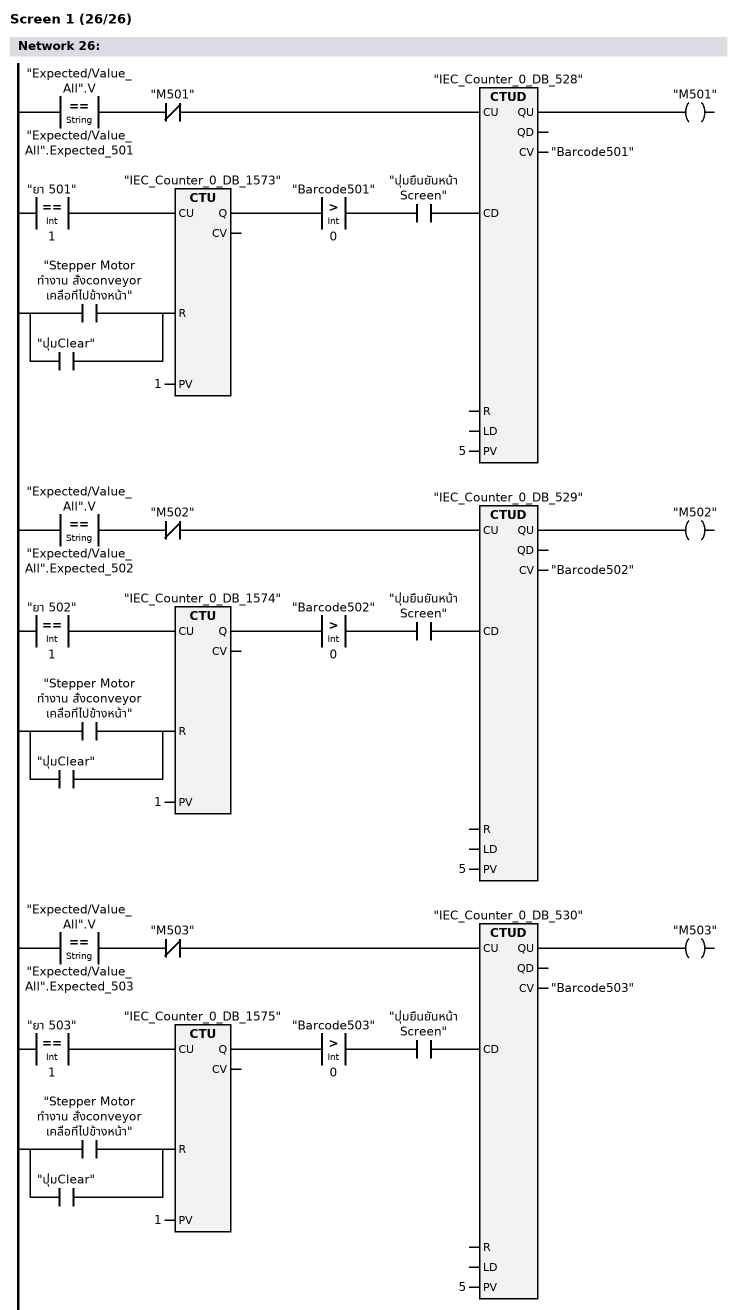
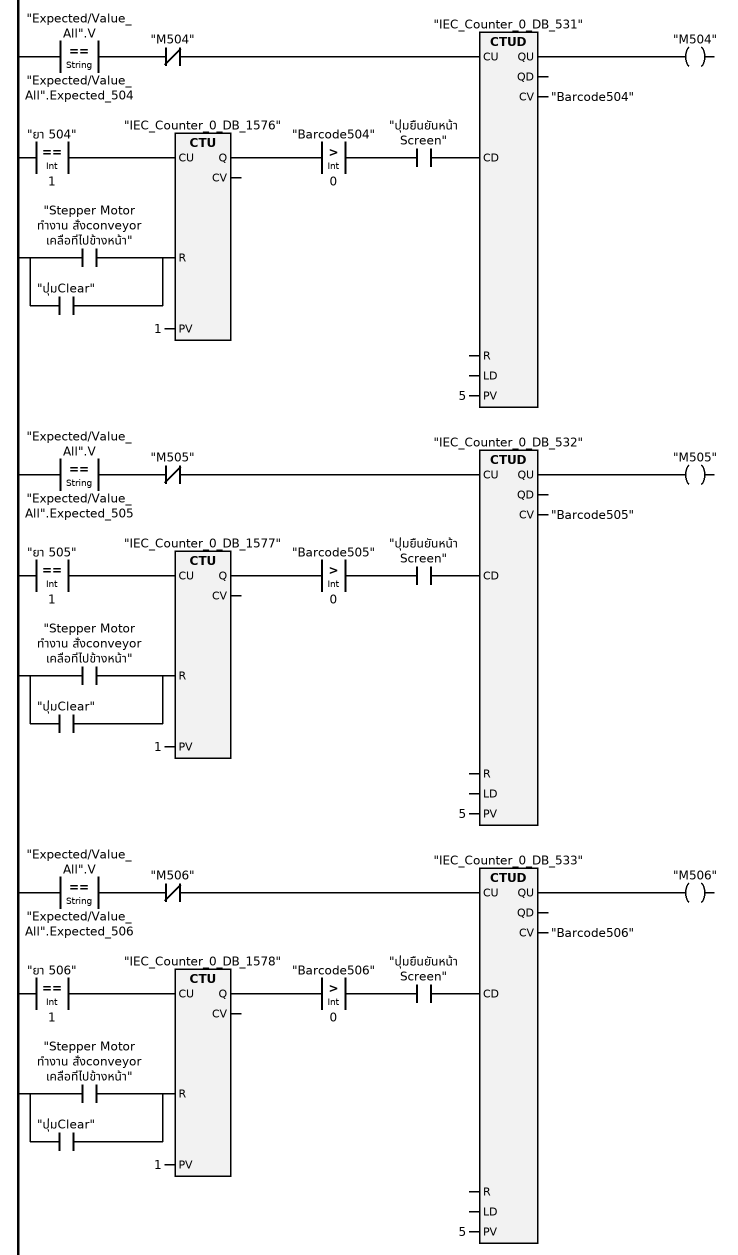
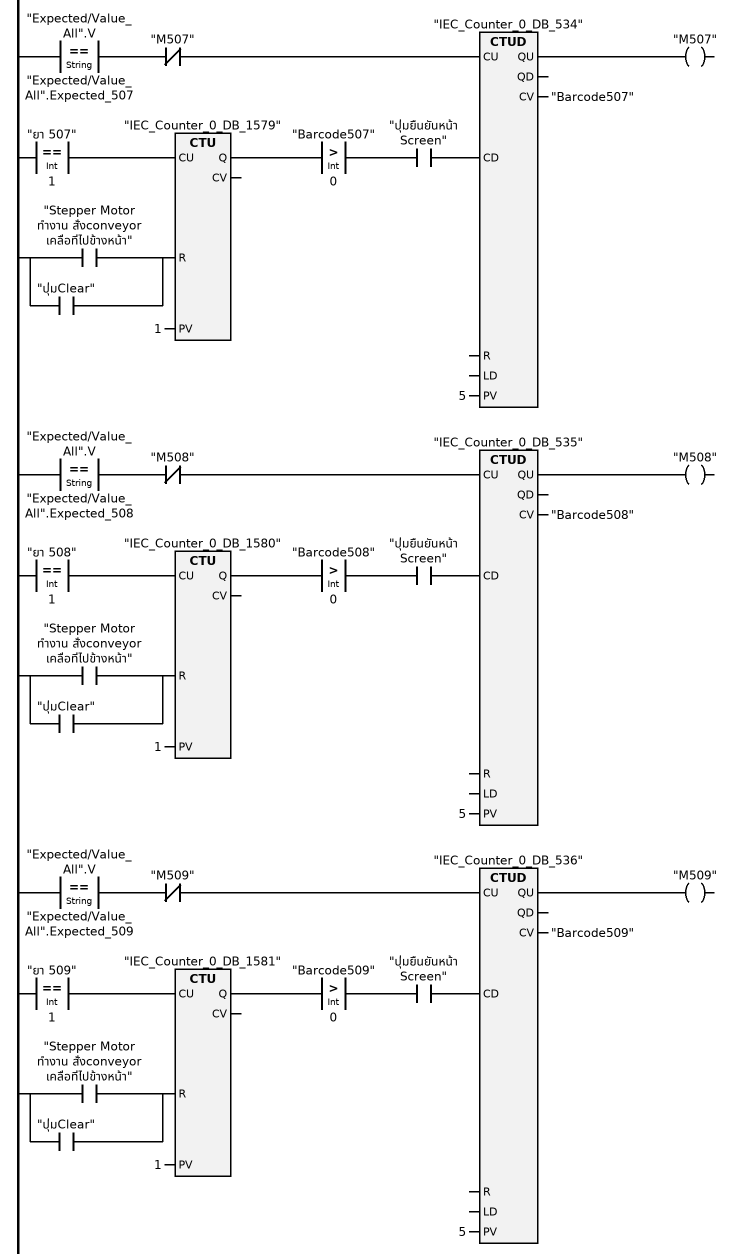
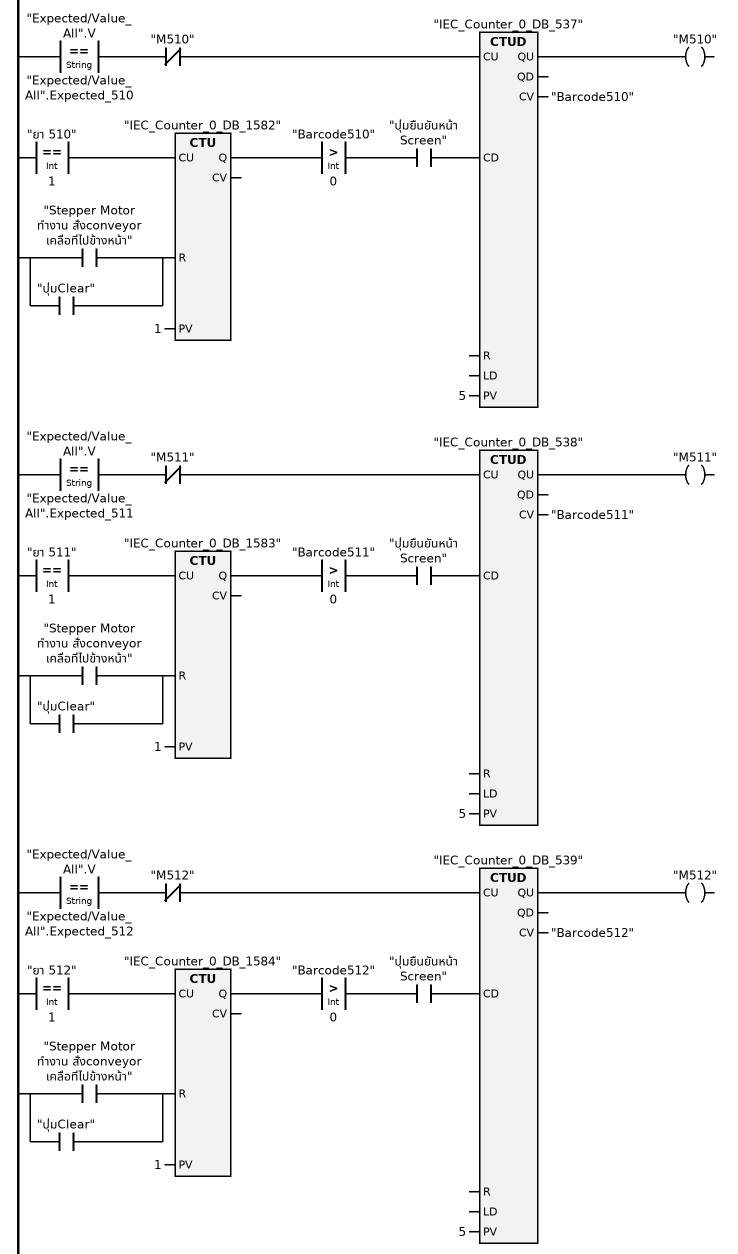
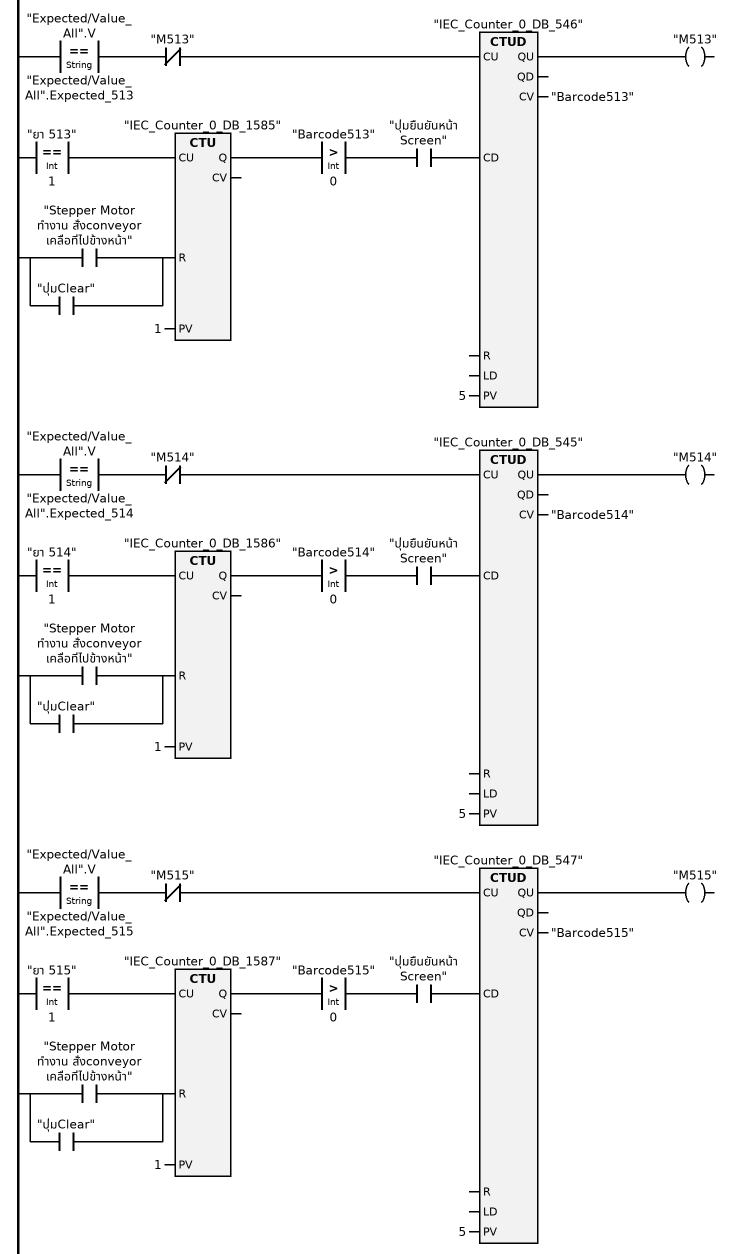
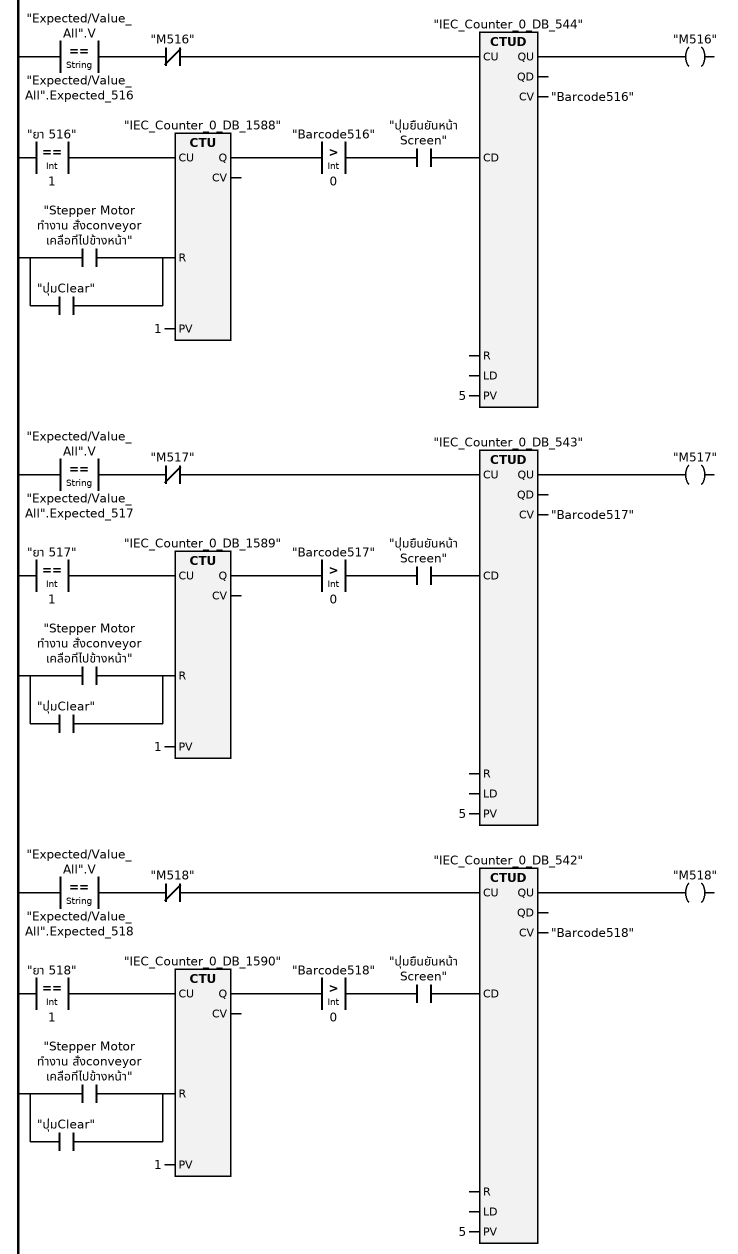
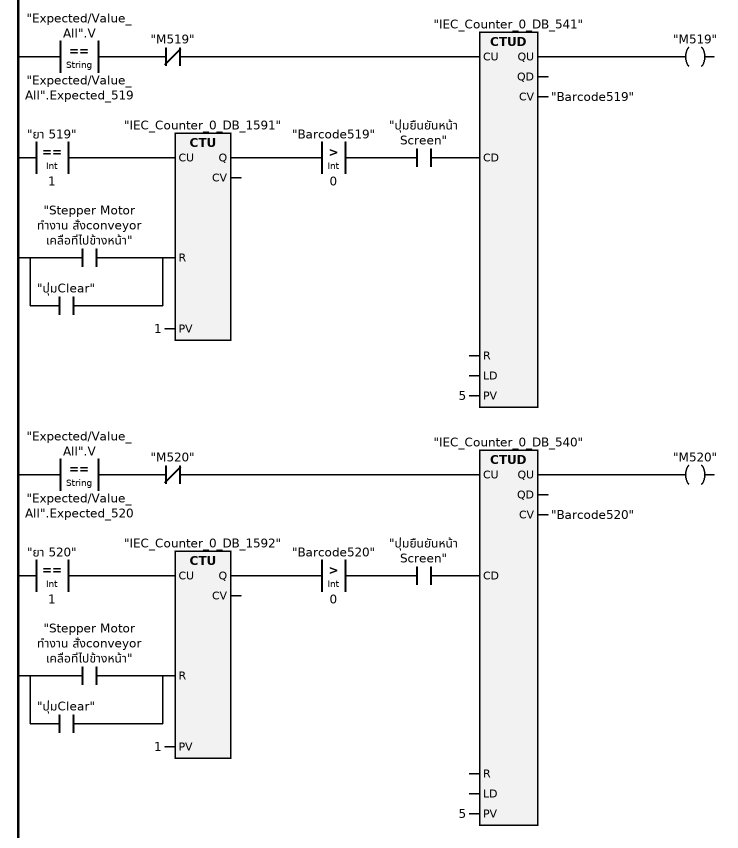
   "IEC_Counter_0_DB_1573".CTU(CU := "ยา 501" = 1,
                           R := "Stepper Motor ทำงาน สั่งconveyor เคลื่อที่ไปข้างหน้า" OR "ปุ่มClear",
                           PV := 1);
   "IEC_Counter_0_DB_528".CTUD(CU := ("Expected/Value_All".V = "Expected/Value_All".Expected_501) AND NOT "M501",
                           CD := "IEC_Counter_0_DB_1573".Q AND ("Barcode501" > 0) AND "ปุ่มยืนยันหน้า Screen",
                           PV := 5,
                           CV => "Barcode501");
   "M501" := "IEC_Counter_0_DB_528".QU;
   "IEC_Counter_0_DB_1574".CTU(CU := "ยา 502" = 1,
                           R := "Stepper Motor ทำงาน สั่งconveyor เคลื่อที่ไปข้างหน้า" OR "ปุ่มClear",
                           PV := 1);
   "IEC_Counter_0_DB_529".CTUD(CU := ("Expected/Value_All".V = "Expected/Value_All".Expected_502) AND NOT "M502",
                           CD := "IEC_Counter_0_DB_1574".Q AND ("Barcode502" > 0) AND "ปุ่มยืนยันหน้า Screen",
                           PV := 5,
                           CV => "Barcode502");
   "M502" := "IEC_Counter_0_DB_529".QU;
   "IEC_Counter_0_DB_1575".CTU(CU := "ยา 503" = 1,
                           R := "Stepper Motor ทำงาน สั่งconveyor เคลื่อที่ไปข้างหน้า" OR "ปุ่มClear",
                           PV := 1);
   "IEC_Counter_0_DB_530".CTUD(CU := ("Expected/Value_All".V = "Expected/Value_All".Expected_503) AND NOT "M503",
                           CD := "IEC_Counter_0_DB_1575".Q AND ("Barcode503" > 0) AND "ปุ่มยืนยันหน้า Screen",
                           PV := 5,
                           CV => "Barcode503");
   "M503" := "IEC_Counter_0_DB_530".QU;
   "IEC_Counter_0_DB_1576".CTU(CU := "ยา 504" = 1,
                           R := "Stepper Motor ทำงาน สั่งconveyor เคลื่อที่ไปข้างหน้า" OR "ปุ่มClear",
                           PV := 1);
   "IEC_Counter_0_DB_531".CTUD(CU := ("Expected/Value_All".V = "Expected/Value_All".Expected_504) AND NOT "M504",
                           CD := "IEC_Counter_0_DB_1576".Q AND ("Barcode504" > 0) AND "ปุ่มยืนยันหน้า Screen",
                           PV := 5,
                           CV => "Barcode504");
   "M504" := "IEC_Counter_0_DB_531".QU;
   "IEC_Counter_0_DB_1577".CTU(CU := "ยา 505" = 1,
                           R := "Stepper Motor ทำงาน สั่งconveyor เคลื่อที่ไปข้างหน้า" OR "ปุ่มClear",
                           PV := 1);
   "IEC_Counter_0_DB_532".CTUD(CU := ("Expected/Value_All".V = "Expected/Value_All".Expected_505) AND NOT "M505",
                           CD := "IEC_Counter_0_DB_1577".Q AND ("Barcode505" > 0) AND "ปุ่มยืนยันหน้า Screen",
                           PV := 5,
                           CV => "Barcode505");
   "M505" := "IEC_Counter_0_DB_532".QU;
   "IEC_Counter_0_DB_1578".CTU(CU := "ยา 506" = 1,
                           R := "Stepper Motor ทำงาน สั่งconveyor เคลื่อที่ไปข้างหน้า" OR "ปุ่มClear",
                           PV := 1);
   "IEC_Counter_0_DB_533".CTUD(CU := ("Expected/Value_All".V = "Expected/Value_All".Expected_506) AND NOT "M506",
                           CD := "IEC_Counter_0_DB_1578".Q AND ("Barcode506" > 0) AND "ปุ่มยืนยันหน้า Screen",
                           PV := 5,
                           CV => "Barcode506");
   "M506" := "IEC_Counter_0_DB_533".QU;
   "IEC_Counter_0_DB_1579".CTU(CU := "ยา 507" = 1,
                           R := "Stepper Motor ทำงาน สั่งconveyor เคลื่อที่ไปข้างหน้า" OR "ปุ่มClear",
                           PV := 1);
   "IEC_Counter_0_DB_534".CTUD(CU := ("Expected/Value_All".V = "Expected/Value_All".Expected_507) AND NOT "M507",
                           CD := "IEC_Counter_0_DB_1579".Q AND ("Barcode507" > 0) AND "ปุ่มยืนยันหน้า Screen",
                           PV := 5,
                           CV => "Barcode507");
   "M507" := "IEC_Counter_0_DB_534".QU;
   "IEC_Counter_0_DB_1580".CTU(CU := "ยา 508" = 1,
                           R := "Stepper Motor ทำงาน สั่งconveyor เคลื่อที่ไปข้างหน้า" OR "ปุ่มClear",
                           PV := 1);
   "IEC_Counter_0_DB_535".CTUD(CU := ("Expected/Value_All".V = "Expected/Value_All".Expected_508) AND NOT "M508",
                           CD := "IEC_Counter_0_DB_1580".Q AND ("Barcode508" > 0) AND "ปุ่มยืนยันหน้า Screen",
                           PV := 5,
                           CV => "Barcode508");
   "M508" := "IEC_Counter_0_DB_535".QU;
   "IEC_Counter_0_DB_1581".CTU(CU := "ยา 509" = 1,
                           R := "Stepper Motor ทำงาน สั่งconveyor เคลื่อที่ไปข้างหน้า" OR "ปุ่มClear",
                           PV := 1);
   "IEC_Counter_0_DB_536".CTUD(CU := ("Expected/Value_All".V = "Expected/Value_All".Expected_509) AND NOT "M509",
                           CD := "IEC_Counter_0_DB_1581".Q AND ("Barcode509" > 0) AND "ปุ่มยืนยันหน้า Screen",
                           PV := 5,
                           CV => "Barcode509");
   "M509" := "IEC_Counter_0_DB_536".QU;
   "IEC_Counter_0_DB_1582".CTU(CU := "ยา 510" = 1,
                           R := "Stepper Motor ทำงาน สั่งconveyor เคลื่อที่ไปข้างหน้า" OR "ปุ่มClear",
                           PV := 1);
   "IEC_Counter_0_DB_537".CTUD(CU := ("Expected/Value_All".V = "Expected/Value_All".Expected_510) AND NOT "M510",
                           CD := "IEC_Counter_0_DB_1582".Q AND ("Barcode510" > 0) AND "ปุ่มยืนยันหน้า Screen",
                           PV := 5,
                           CV => "Barcode510");
   "M510" := "IEC_Counter_0_DB_537".QU;
   "IEC_Counter_0_DB_1583".CTU(CU := "ยา 511" = 1,
                           R := "Stepper Motor ทำงาน สั่งconveyor เคลื่อที่ไปข้างหน้า" OR "ปุ่มClear",
                           PV := 1);
   "IEC_Counter_0_DB_538".CTUD(CU := ("Expected/Value_All".V = "Expected/Value_All".Expected_511) AND NOT "M511",
                           CD := "IEC_Counter_0_DB_1583".Q AND ("Barcode511" > 0) AND "ปุ่มยืนยันหน้า Screen",
                           PV := 5,
                           CV => "Barcode511");
   "M511" := "IEC_Counter_0_DB_538".QU;
   "IEC_Counter_0_DB_1584".CTU(CU := "ยา 512" = 1,
                           R := "Stepper Motor ทำงาน สั่งconveyor เคลื่อที่ไปข้างหน้า" OR "ปุ่มClear",
                           PV := 1);
   "IEC_Counter_0_DB_539".CTUD(CU := ("Expected/Value_All".V = "Expected/Value_All".Expected_512) AND NOT "M512",
                           CD := "IEC_Counter_0_DB_1584".Q AND ("Barcode512" > 0) AND "ปุ่มยืนยันหน้า Screen",
                           PV := 5,
                           CV => "Barcode512");
   "M512" := "IEC_Counter_0_DB_539".QU;
   "IEC_Counter_0_DB_1585".CTU(CU := "ยา 513" = 1,
                           R := "Stepper Motor ทำงาน สั่งconveyor เคลื่อที่ไปข้างหน้า" OR "ปุ่มClear",
                           PV := 1);
   "IEC_Counter_0_DB_546".CTUD(CU := ("Expected/Value_All".V = "Expected/Value_All".Expected_513) AND NOT "M513",
                           CD := "IEC_Counter_0_DB_1585".Q AND ("Barcode513" > 0) AND "ปุ่มยืนยันหน้า Screen",
                           PV := 5,
                           CV => "Barcode513");
   "M513" := "IEC_Counter_0_DB_546".QU;
   "IEC_Counter_0_DB_1586".CTU(CU := "ยา 514" = 1,
                           R := "Stepper Motor ทำงาน สั่งconveyor เคลื่อที่ไปข้างหน้า" OR "ปุ่มClear",
                           PV := 1);
   "IEC_Counter_0_DB_545".CTUD(CU := ("Expected/Value_All".V = "Expected/Value_All".Expected_514) AND NOT "M514",
                           CD := "IEC_Counter_0_DB_1586".Q AND ("Barcode514" > 0) AND "ปุ่มยืนยันหน้า Screen",
                           PV := 5,
                           CV => "Barcode514");
   "M514" := "IEC_Counter_0_DB_545".QU;
   "IEC_Counter_0_DB_1587".CTU(CU := "ยา 515" = 1,
                           R := "Stepper Motor ทำงาน สั่งconveyor เคลื่อที่ไปข้างหน้า" OR "ปุ่มClear",
                           PV := 1);
   "IEC_Counter_0_DB_547".CTUD(CU := ("Expected/Value_All".V = "Expected/Value_All".Expected_515) AND NOT "M515",
                           CD := "IEC_Counter_0_DB_1587".Q AND ("Barcode515" > 0) AND "ปุ่มยืนยันหน้า Screen",
                           PV := 5,
                           CV => "Barcode515");
   "M515" := "IEC_Counter_0_DB_547".QU;
   "IEC_Counter_0_DB_1588".CTU(CU := "ยา 516" = 1,
                           R := "Stepper Motor ทำงาน สั่งconveyor เคลื่อที่ไปข้างหน้า" OR "ปุ่มClear",
                           PV := 1);
   "IEC_Counter_0_DB_544".CTUD(CU := ("Expected/Value_All".V = "Expected/Value_All".Expected_516) AND NOT "M516",
                           CD := "IEC_Counter_0_DB_1588".Q AND ("Barcode516" > 0) AND "ปุ่มยืนยันหน้า Screen",
                           PV := 5,
                           CV => "Barcode516");
   "M516" := "IEC_Counter_0_DB_544".QU;
   "IEC_Counter_0_DB_1589".CTU(CU := "ยา 517" = 1,
                           R := "Stepper Motor ทำงาน สั่งconveyor เคลื่อที่ไปข้างหน้า" OR "ปุ่มClear",
                           PV := 1);
   "IEC_Counter_0_DB_543".CTUD(CU := ("Expected/Value_All".V = "Expected/Value_All".Expected_517) AND NOT "M517",
                           CD := "IEC_Counter_0_DB_1589".Q AND ("Barcode517" > 0) AND "ปุ่มยืนยันหน้า Screen",
                           PV := 5,
                           CV => "Barcode517");
   "M517" := "IEC_Counter_0_DB_543".QU;
   "IEC_Counter_0_DB_1590".CTU(CU := "ยา 518" = 1,
                           R := "Stepper Motor ทำงาน สั่งconveyor เคลื่อที่ไปข้างหน้า" OR "ปุ่มClear",
                           PV := 1);
   "IEC_Counter_0_DB_542".CTUD(CU := ("Expected/Value_All".V = "Expected/Value_All".Expected_518) AND NOT "M518",
                           CD := "IEC_Counter_0_DB_1590".Q AND ("Barcode518" > 0) AND "ปุ่มยืนยันหน้า Screen",
                           PV := 5,
                           CV => "Barcode518");
   "M518" := "IEC_Counter_0_DB_542".QU;
   "IEC_Counter_0_DB_1591".CTU(CU := "ยา 519" = 1,
                           R := "Stepper Motor ทำงาน สั่งconveyor เคลื่อที่ไปข้างหน้า" OR "ปุ่มClear",
                           PV := 1);
   "IEC_Counter_0_DB_541".CTUD(CU := ("Expected/Value_All".V = "Expected/Value_All".Expected_519) AND NOT "M519",
                           CD := "IEC_Counter_0_DB_1591".Q AND ("Barcode519" > 0) AND "ปุ่มยืนยันหน้า Screen",
                           PV := 5,
                           CV => "Barcode519");
   "M519" := "IEC_Counter_0_DB_541".QU;
   "IEC_Counter_0_DB_1592".CTU(CU := "ยา 520" = 1,
                           R := "Stepper Motor ทำงาน สั่งconveyor เคลื่อที่ไปข้างหน้า" OR "ปุ่มClear",
                           PV := 1);
   "IEC_Counter_0_DB_540".CTUD(CU := ("Expected/Value_All".V = "Expected/Value_All".Expected_520) AND NOT "M520",
                           CD := "IEC_Counter_0_DB_1592".Q AND ("Barcode520" > 0) AND "ปุ่มยืนยันหน้า Screen",
                           PV := 5,
                           CV => "Barcode520");
   "M520" := "IEC_Counter_0_DB_540".QU;
END_REGION
END_FUNCTION

FUNCTION "Screen2" : Void   // FC14, LAD
{ S7_Optimized_Access := 'TRUE' }
VERSION : 0.1
   VAR_OUTPUT
      Output : Word;
   END_VAR
BEGIN

REGION Network 1
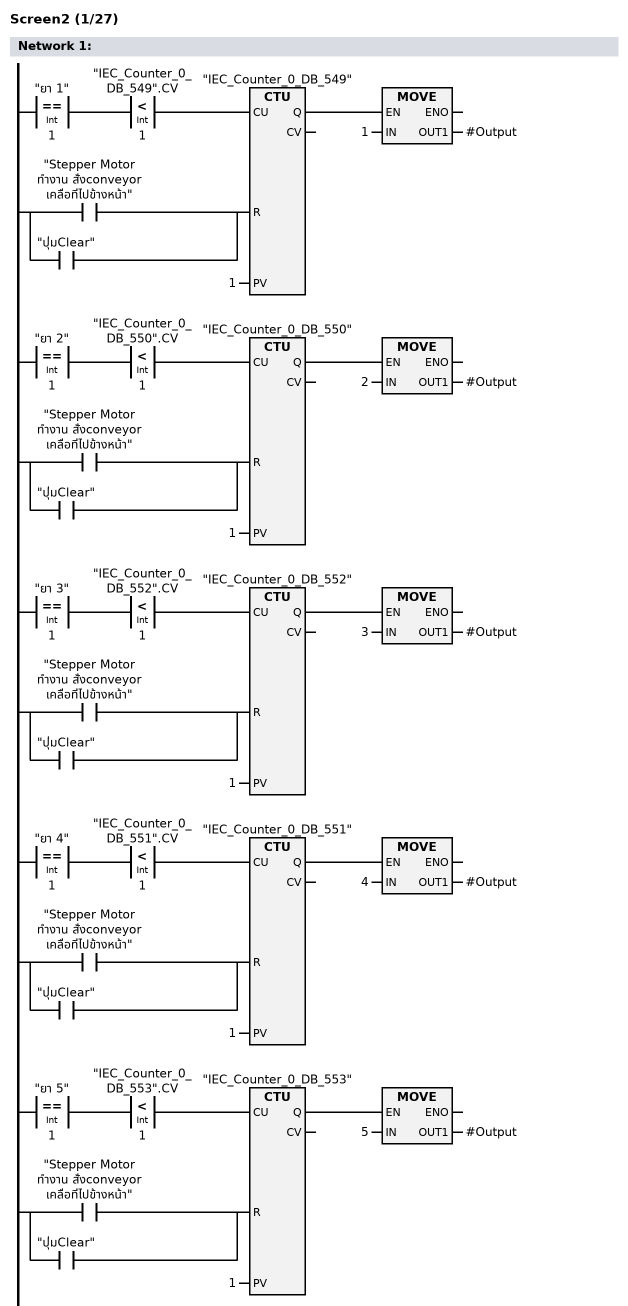
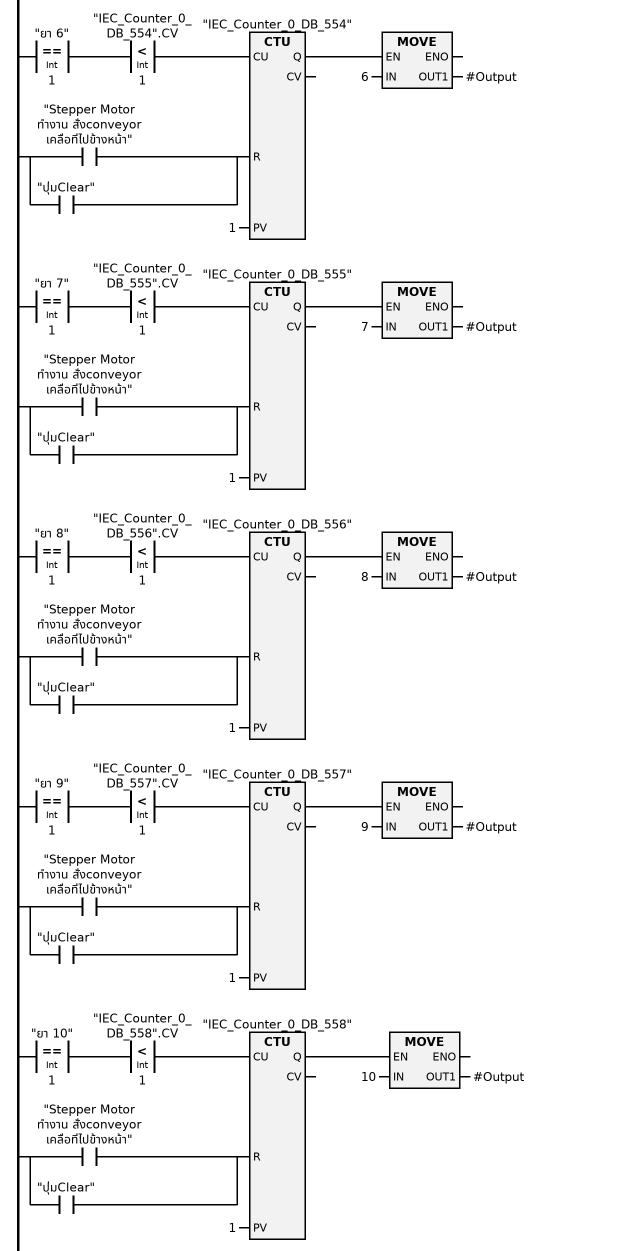
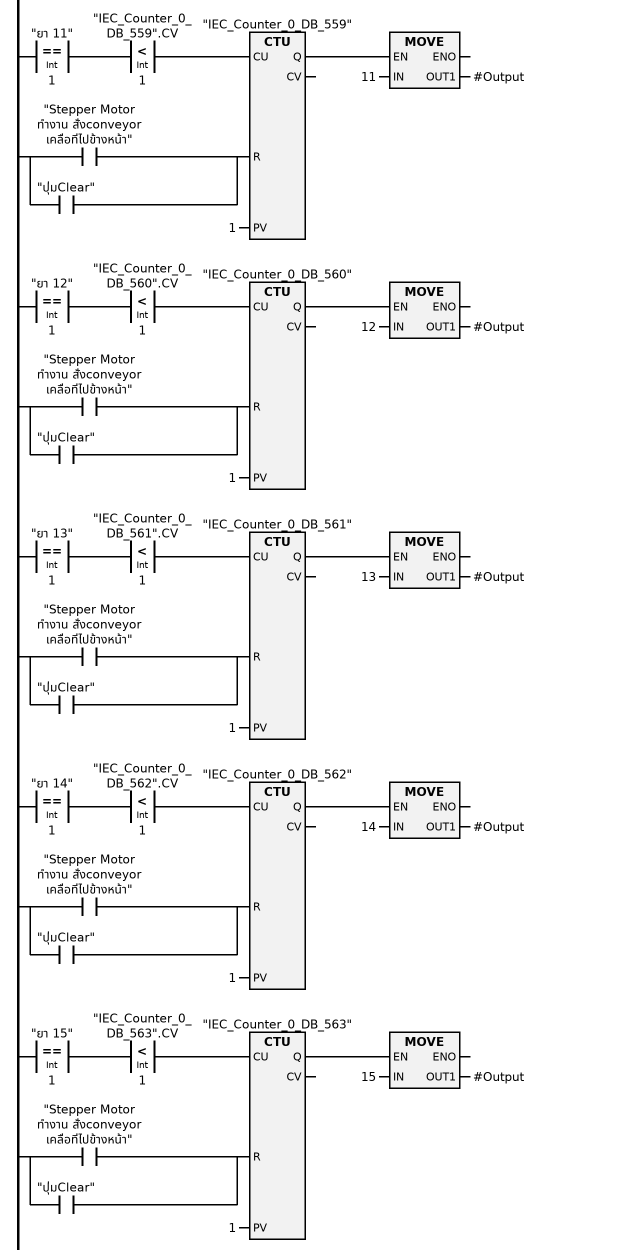
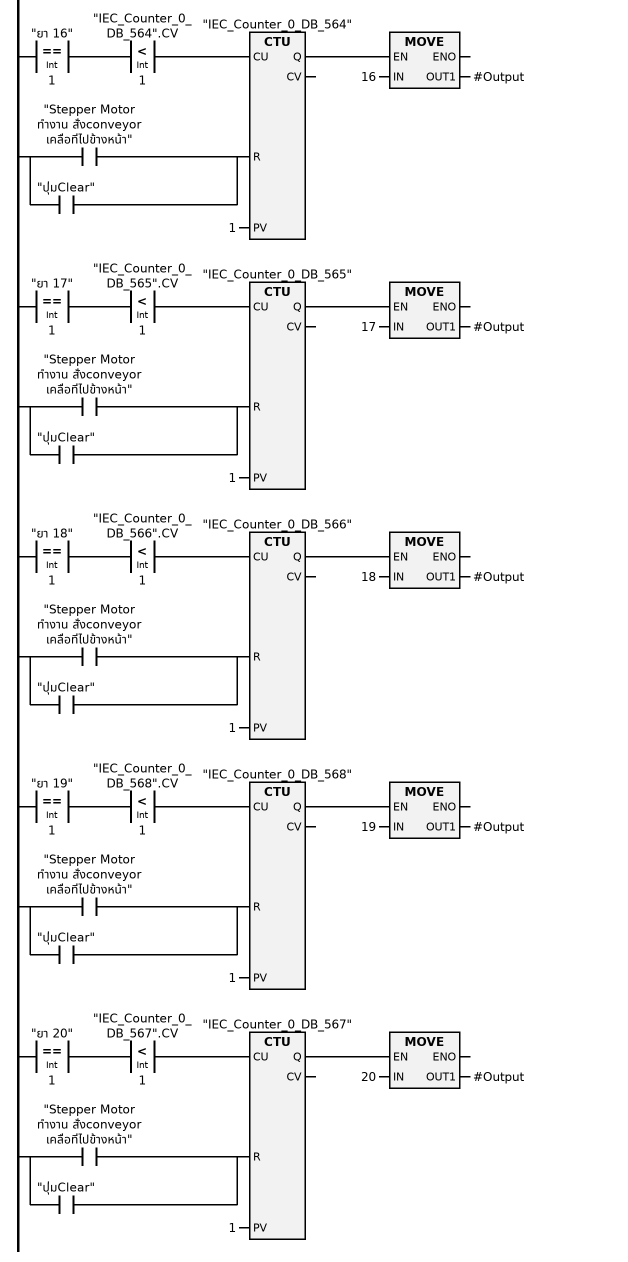
   "IEC_Counter_0_DB_549".CTU(CU := ("ยา 1" = 1) AND ("IEC_Counter_0_DB_549".CV < 1),
                           R := "Stepper Motor ทำงาน สั่งconveyor เคลื่อที่ไปข้างหน้า" OR "ปุ่มClear",
                           PV := 1);
   IF "IEC_Counter_0_DB_549".Q THEN #Output := 1; END_IF;
   "IEC_Counter_0_DB_550".CTU(CU := ("ยา 2" = 1) AND ("IEC_Counter_0_DB_550".CV < 1),
                           R := "Stepper Motor ทำงาน สั่งconveyor เคลื่อที่ไปข้างหน้า" OR "ปุ่มClear",
                           PV := 1);
   IF "IEC_Counter_0_DB_550".Q THEN #Output := 2; END_IF;
   "IEC_Counter_0_DB_552".CTU(CU := ("ยา 3" = 1) AND ("IEC_Counter_0_DB_552".CV < 1),
                           R := "Stepper Motor ทำงาน สั่งconveyor เคลื่อที่ไปข้างหน้า" OR "ปุ่มClear",
                           PV := 1);
   IF "IEC_Counter_0_DB_552".Q THEN #Output := 3; END_IF;
   "IEC_Counter_0_DB_551".CTU(CU := ("ยา 4" = 1) AND ("IEC_Counter_0_DB_551".CV < 1),
                           R := "Stepper Motor ทำงาน สั่งconveyor เคลื่อที่ไปข้างหน้า" OR "ปุ่มClear",
                           PV := 1);
   IF "IEC_Counter_0_DB_551".Q THEN #Output := 4; END_IF;
   "IEC_Counter_0_DB_553".CTU(CU := ("ยา 5" = 1) AND ("IEC_Counter_0_DB_553".CV < 1),
                           R := "Stepper Motor ทำงาน สั่งconveyor เคลื่อที่ไปข้างหน้า" OR "ปุ่มClear",
                           PV := 1);
   IF "IEC_Counter_0_DB_553".Q THEN #Output := 5; END_IF;
   "IEC_Counter_0_DB_554".CTU(CU := ("ยา 6" = 1) AND ("IEC_Counter_0_DB_554".CV < 1),
                           R := "Stepper Motor ทำงาน สั่งconveyor เคลื่อที่ไปข้างหน้า" OR "ปุ่มClear",
                           PV := 1);
   IF "IEC_Counter_0_DB_554".Q THEN #Output := 6; END_IF;
   "IEC_Counter_0_DB_555".CTU(CU := ("ยา 7" = 1) AND ("IEC_Counter_0_DB_555".CV < 1),
                           R := "Stepper Motor ทำงาน สั่งconveyor เคลื่อที่ไปข้างหน้า" OR "ปุ่มClear",
                           PV := 1);
   IF "IEC_Counter_0_DB_555".Q THEN #Output := 7; END_IF;
   "IEC_Counter_0_DB_556".CTU(CU := ("ยา 8" = 1) AND ("IEC_Counter_0_DB_556".CV < 1),
                           R := "Stepper Motor ทำงาน สั่งconveyor เคลื่อที่ไปข้างหน้า" OR "ปุ่มClear",
                           PV := 1);
   IF "IEC_Counter_0_DB_556".Q THEN #Output := 8; END_IF;
   "IEC_Counter_0_DB_557".CTU(CU := ("ยา 9" = 1) AND ("IEC_Counter_0_DB_557".CV < 1),
                           R := "Stepper Motor ทำงาน สั่งconveyor เคลื่อที่ไปข้างหน้า" OR "ปุ่มClear",
                           PV := 1);
   IF "IEC_Counter_0_DB_557".Q THEN #Output := 9; END_IF;
   "IEC_Counter_0_DB_558".CTU(CU := ("ยา 10" = 1) AND ("IEC_Counter_0_DB_558".CV < 1),
                           R := "Stepper Motor ทำงาน สั่งconveyor เคลื่อที่ไปข้างหน้า" OR "ปุ่มClear",
                           PV := 1);
   IF "IEC_Counter_0_DB_558".Q THEN #Output := 10; END_IF;
   "IEC_Counter_0_DB_559".CTU(CU := ("ยา 11" = 1) AND ("IEC_Counter_0_DB_559".CV < 1),
                           R := "Stepper Motor ทำงาน สั่งconveyor เคลื่อที่ไปข้างหน้า" OR "ปุ่มClear",
                           PV := 1);
   IF "IEC_Counter_0_DB_559".Q THEN #Output := 11; END_IF;
   "IEC_Counter_0_DB_560".CTU(CU := ("ยา 12" = 1) AND ("IEC_Counter_0_DB_560".CV < 1),
                           R := "Stepper Motor ทำงาน สั่งconveyor เคลื่อที่ไปข้างหน้า" OR "ปุ่มClear",
                           PV := 1);
   IF "IEC_Counter_0_DB_560".Q THEN #Output := 12; END_IF;
   "IEC_Counter_0_DB_561".CTU(CU := ("ยา 13" = 1) AND ("IEC_Counter_0_DB_561".CV < 1),
                           R := "Stepper Motor ทำงาน สั่งconveyor เคลื่อที่ไปข้างหน้า" OR "ปุ่มClear",
                           PV := 1);
   IF "IEC_Counter_0_DB_561".Q THEN #Output := 13; END_IF;
   "IEC_Counter_0_DB_562".CTU(CU := ("ยา 14" = 1) AND ("IEC_Counter_0_DB_562".CV < 1),
                           R := "Stepper Motor ทำงาน สั่งconveyor เคลื่อที่ไปข้างหน้า" OR "ปุ่มClear",
                           PV := 1);
   IF "IEC_Counter_0_DB_562".Q THEN #Output := 14; END_IF;
   "IEC_Counter_0_DB_563".CTU(CU := ("ยา 15" = 1) AND ("IEC_Counter_0_DB_563".CV < 1),
                           R := "Stepper Motor ทำงาน สั่งconveyor เคลื่อที่ไปข้างหน้า" OR "ปุ่มClear",
                           PV := 1);
   IF "IEC_Counter_0_DB_563".Q THEN #Output := 15; END_IF;
   "IEC_Counter_0_DB_564".CTU(CU := ("ยา 16" = 1) AND ("IEC_Counter_0_DB_564".CV < 1),
                           R := "Stepper Motor ทำงาน สั่งconveyor เคลื่อที่ไปข้างหน้า" OR "ปุ่มClear",
                           PV := 1);
   IF "IEC_Counter_0_DB_564".Q THEN #Output := 16; END_IF;
   "IEC_Counter_0_DB_565".CTU(CU := ("ยา 17" = 1) AND ("IEC_Counter_0_DB_565".CV < 1),
                           R := "Stepper Motor ทำงาน สั่งconveyor เคลื่อที่ไปข้างหน้า" OR "ปุ่มClear",
                           PV := 1);
   IF "IEC_Counter_0_DB_565".Q THEN #Output := 17; END_IF;
   "IEC_Counter_0_DB_566".CTU(CU := ("ยา 18" = 1) AND ("IEC_Counter_0_DB_566".CV < 1),
                           R := "Stepper Motor ทำงาน สั่งconveyor เคลื่อที่ไปข้างหน้า" OR "ปุ่มClear",
                           PV := 1);
   IF "IEC_Counter_0_DB_566".Q THEN #Output := 18; END_IF;
   "IEC_Counter_0_DB_568".CTU(CU := ("ยา 19" = 1) AND ("IEC_Counter_0_DB_568".CV < 1),
                           R := "Stepper Motor ทำงาน สั่งconveyor เคลื่อที่ไปข้างหน้า" OR "ปุ่มClear",
                           PV := 1);
   IF "IEC_Counter_0_DB_568".Q THEN #Output := 19; END_IF;
   "IEC_Counter_0_DB_567".CTU(CU := ("ยา 20" = 1) AND ("IEC_Counter_0_DB_567".CV < 1),
                           R := "Stepper Motor ทำงาน สั่งconveyor เคลื่อที่ไปข้างหน้า" OR "ปุ่มClear",
                           PV := 1);
   IF "IEC_Counter_0_DB_567".Q THEN #Output := 20; END_IF;
END_REGION

REGION Network 2
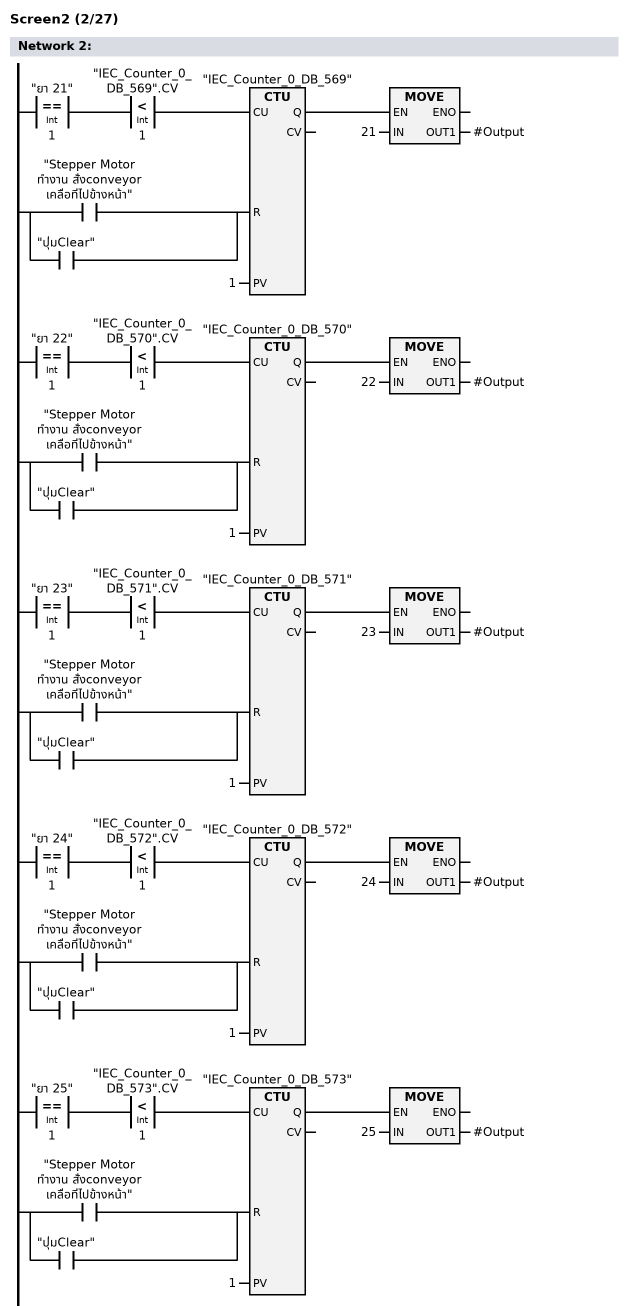
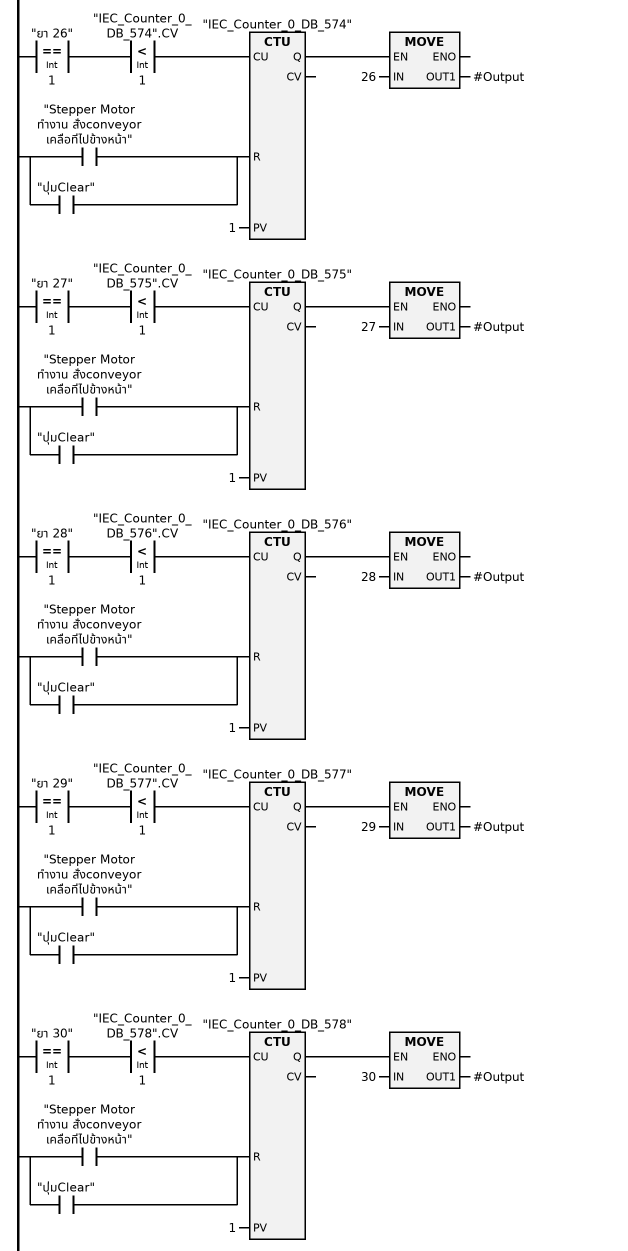
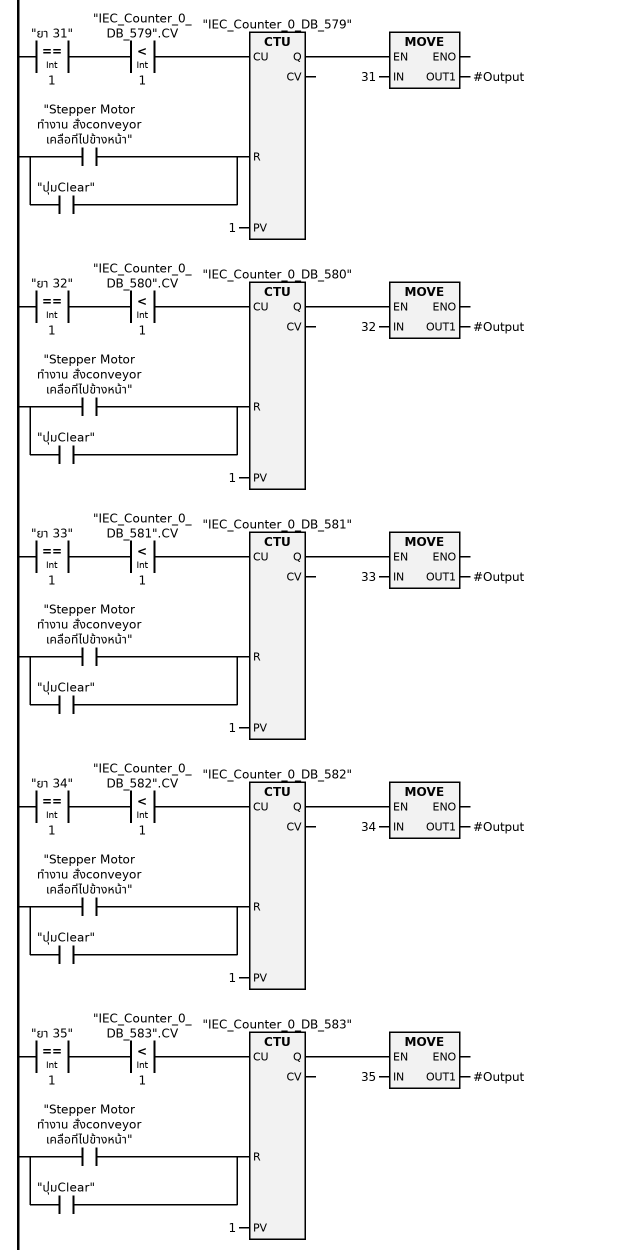
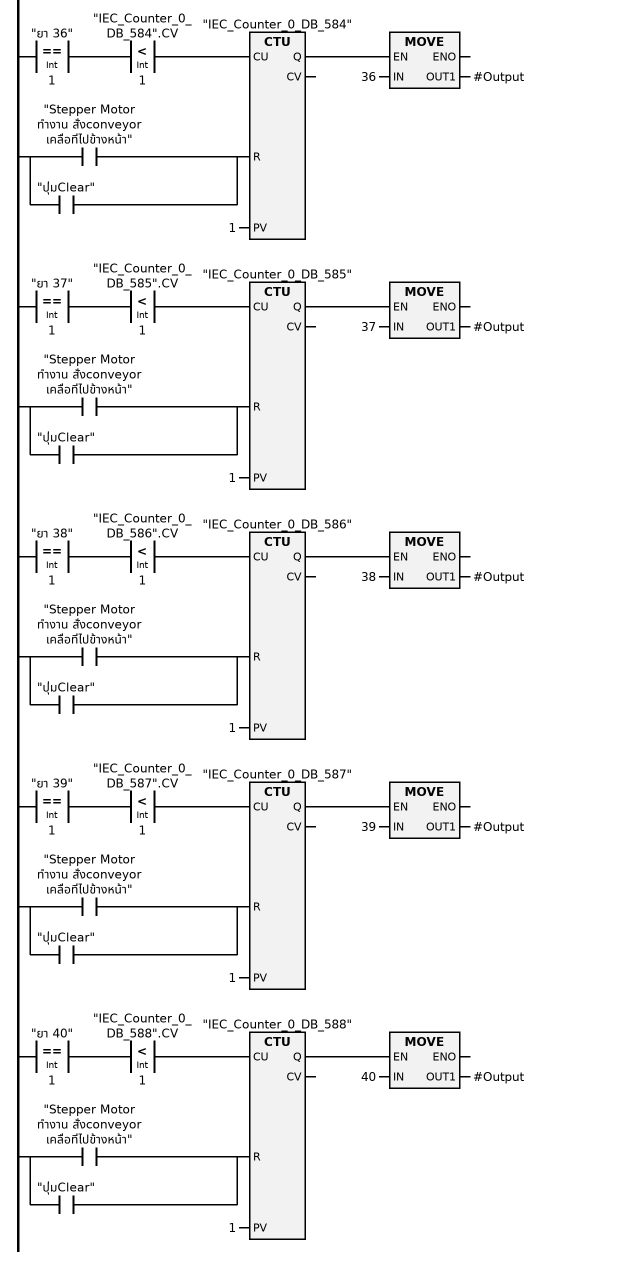
   "IEC_Counter_0_DB_569".CTU(CU := ("ยา 21" = 1) AND ("IEC_Counter_0_DB_569".CV < 1),
                           R := "Stepper Motor ทำงาน สั่งconveyor เคลื่อที่ไปข้างหน้า" OR "ปุ่มClear",
                           PV := 1);
   IF "IEC_Counter_0_DB_569".Q THEN #Output := 21; END_IF;
   "IEC_Counter_0_DB_570".CTU(CU := ("ยา 22" = 1) AND ("IEC_Counter_0_DB_570".CV < 1),
                           R := "Stepper Motor ทำงาน สั่งconveyor เคลื่อที่ไปข้างหน้า" OR "ปุ่มClear",
                           PV := 1);
   IF "IEC_Counter_0_DB_570".Q THEN #Output := 22; END_IF;
   "IEC_Counter_0_DB_571".CTU(CU := ("ยา 23" = 1) AND ("IEC_Counter_0_DB_571".CV < 1),
                           R := "Stepper Motor ทำงาน สั่งconveyor เคลื่อที่ไปข้างหน้า" OR "ปุ่มClear",
                           PV := 1);
   IF "IEC_Counter_0_DB_571".Q THEN #Output := 23; END_IF;
   "IEC_Counter_0_DB_572".CTU(CU := ("ยา 24" = 1) AND ("IEC_Counter_0_DB_572".CV < 1),
                           R := "Stepper Motor ทำงาน สั่งconveyor เคลื่อที่ไปข้างหน้า" OR "ปุ่มClear",
                           PV := 1);
   IF "IEC_Counter_0_DB_572".Q THEN #Output := 24; END_IF;
   "IEC_Counter_0_DB_573".CTU(CU := ("ยา 25" = 1) AND ("IEC_Counter_0_DB_573".CV < 1),
                           R := "Stepper Motor ทำงาน สั่งconveyor เคลื่อที่ไปข้างหน้า" OR "ปุ่มClear",
                           PV := 1);
   IF "IEC_Counter_0_DB_573".Q THEN #Output := 25; END_IF;
   "IEC_Counter_0_DB_574".CTU(CU := ("ยา 26" = 1) AND ("IEC_Counter_0_DB_574".CV < 1),
                           R := "Stepper Motor ทำงาน สั่งconveyor เคลื่อที่ไปข้างหน้า" OR "ปุ่มClear",
                           PV := 1);
   IF "IEC_Counter_0_DB_574".Q THEN #Output := 26; END_IF;
   "IEC_Counter_0_DB_575".CTU(CU := ("ยา 27" = 1) AND ("IEC_Counter_0_DB_575".CV < 1),
                           R := "Stepper Motor ทำงาน สั่งconveyor เคลื่อที่ไปข้างหน้า" OR "ปุ่มClear",
                           PV := 1);
   IF "IEC_Counter_0_DB_575".Q THEN #Output := 27; END_IF;
   "IEC_Counter_0_DB_576".CTU(CU := ("ยา 28" = 1) AND ("IEC_Counter_0_DB_576".CV < 1),
                           R := "Stepper Motor ทำงาน สั่งconveyor เคลื่อที่ไปข้างหน้า" OR "ปุ่มClear",
                           PV := 1);
   IF "IEC_Counter_0_DB_576".Q THEN #Output := 28; END_IF;
   "IEC_Counter_0_DB_577".CTU(CU := ("ยา 29" = 1) AND ("IEC_Counter_0_DB_577".CV < 1),
                           R := "Stepper Motor ทำงาน สั่งconveyor เคลื่อที่ไปข้างหน้า" OR "ปุ่มClear",
                           PV := 1);
   IF "IEC_Counter_0_DB_577".Q THEN #Output := 29; END_IF;
   "IEC_Counter_0_DB_578".CTU(CU := ("ยา 30" = 1) AND ("IEC_Counter_0_DB_578".CV < 1),
                           R := "Stepper Motor ทำงาน สั่งconveyor เคลื่อที่ไปข้างหน้า" OR "ปุ่มClear",
                           PV := 1);
   IF "IEC_Counter_0_DB_578".Q THEN #Output := 30; END_IF;
   "IEC_Counter_0_DB_579".CTU(CU := ("ยา 31" = 1) AND ("IEC_Counter_0_DB_579".CV < 1),
                           R := "Stepper Motor ทำงาน สั่งconveyor เคลื่อที่ไปข้างหน้า" OR "ปุ่มClear",
                           PV := 1);
   IF "IEC_Counter_0_DB_579".Q THEN #Output := 31; END_IF;
   "IEC_Counter_0_DB_580".CTU(CU := ("ยา 32" = 1) AND ("IEC_Counter_0_DB_580".CV < 1),
                           R := "Stepper Motor ทำงาน สั่งconveyor เคลื่อที่ไปข้างหน้า" OR "ปุ่มClear",
                           PV := 1);
   IF "IEC_Counter_0_DB_580".Q THEN #Output := 32; END_IF;
   "IEC_Counter_0_DB_581".CTU(CU := ("ยา 33" = 1) AND ("IEC_Counter_0_DB_581".CV < 1),
                           R := "Stepper Motor ทำงาน สั่งconveyor เคลื่อที่ไปข้างหน้า" OR "ปุ่มClear",
                           PV := 1);
   IF "IEC_Counter_0_DB_581".Q THEN #Output := 33; END_IF;
   "IEC_Counter_0_DB_582".CTU(CU := ("ยา 34" = 1) AND ("IEC_Counter_0_DB_582".CV < 1),
                           R := "Stepper Motor ทำงาน สั่งconveyor เคลื่อที่ไปข้างหน้า" OR "ปุ่มClear",
                           PV := 1);
   IF "IEC_Counter_0_DB_582".Q THEN #Output := 34; END_IF;
   "IEC_Counter_0_DB_583".CTU(CU := ("ยา 35" = 1) AND ("IEC_Counter_0_DB_583".CV < 1),
                           R := "Stepper Motor ทำงาน สั่งconveyor เคลื่อที่ไปข้างหน้า" OR "ปุ่มClear",
                           PV := 1);
   IF "IEC_Counter_0_DB_583".Q THEN #Output := 35; END_IF;
   "IEC_Counter_0_DB_584".CTU(CU := ("ยา 36" = 1) AND ("IEC_Counter_0_DB_584".CV < 1),
                           R := "Stepper Motor ทำงาน สั่งconveyor เคลื่อที่ไปข้างหน้า" OR "ปุ่มClear",
                           PV := 1);
   IF "IEC_Counter_0_DB_584".Q THEN #Output := 36; END_IF;
   "IEC_Counter_0_DB_585".CTU(CU := ("ยา 37" = 1) AND ("IEC_Counter_0_DB_585".CV < 1),
                           R := "Stepper Motor ทำงาน สั่งconveyor เคลื่อที่ไปข้างหน้า" OR "ปุ่มClear",
                           PV := 1);
   IF "IEC_Counter_0_DB_585".Q THEN #Output := 37; END_IF;
   "IEC_Counter_0_DB_586".CTU(CU := ("ยา 38" = 1) AND ("IEC_Counter_0_DB_586".CV < 1),
                           R := "Stepper Motor ทำงาน สั่งconveyor เคลื่อที่ไปข้างหน้า" OR "ปุ่มClear",
                           PV := 1);
   IF "IEC_Counter_0_DB_586".Q THEN #Output := 38; END_IF;
   "IEC_Counter_0_DB_587".CTU(CU := ("ยา 39" = 1) AND ("IEC_Counter_0_DB_587".CV < 1),
                           R := "Stepper Motor ทำงาน สั่งconveyor เคลื่อที่ไปข้างหน้า" OR "ปุ่มClear",
                           PV := 1);
   IF "IEC_Counter_0_DB_587".Q THEN #Output := 39; END_IF;
   "IEC_Counter_0_DB_588".CTU(CU := ("ยา 40" = 1) AND ("IEC_Counter_0_DB_588".CV < 1),
                           R := "Stepper Motor ทำงาน สั่งconveyor เคลื่อที่ไปข้างหน้า" OR "ปุ่มClear",
                           PV := 1);
   IF "IEC_Counter_0_DB_588".Q THEN #Output := 40; END_IF;
END_REGION

REGION Network 3
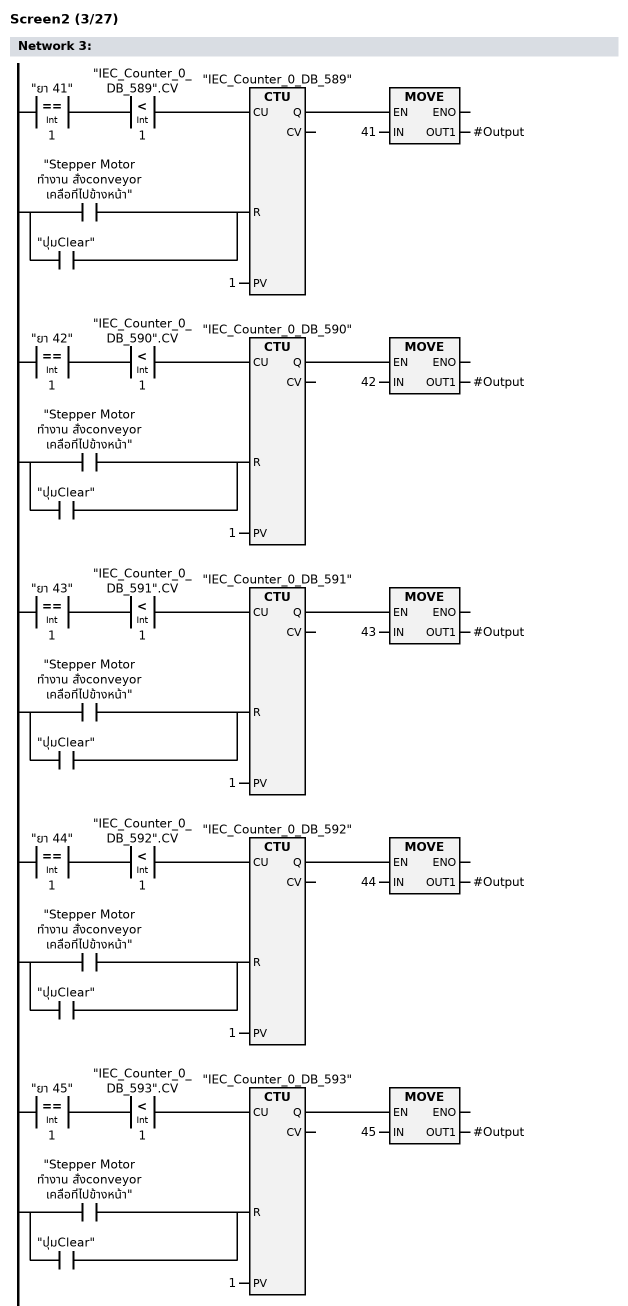
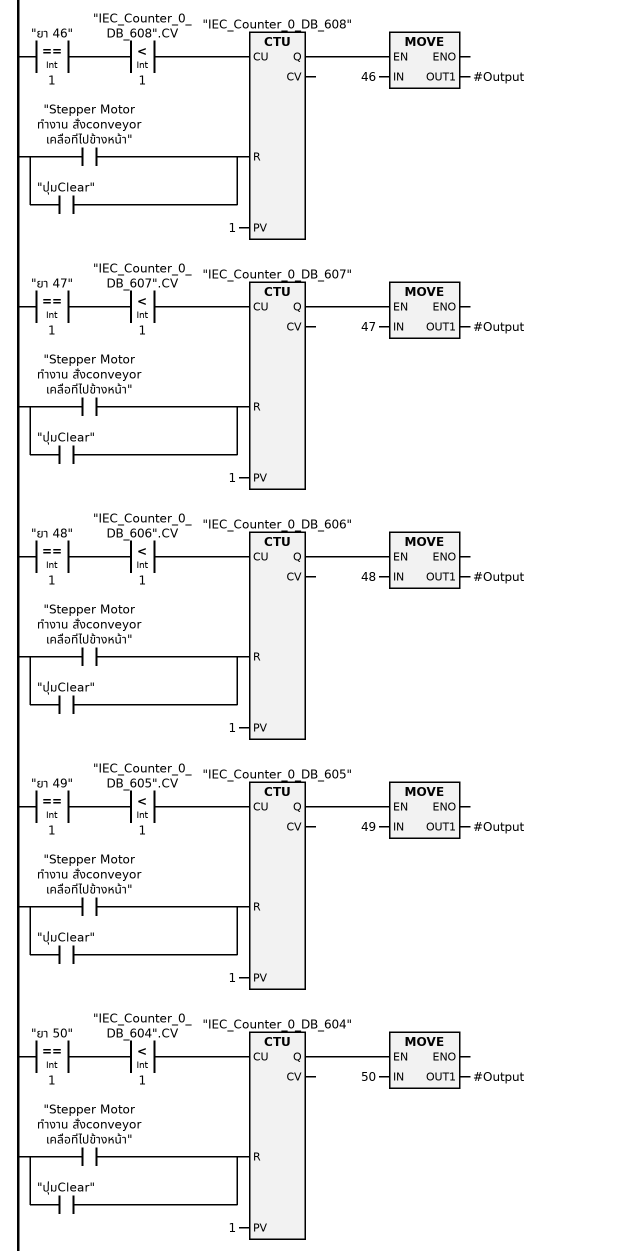
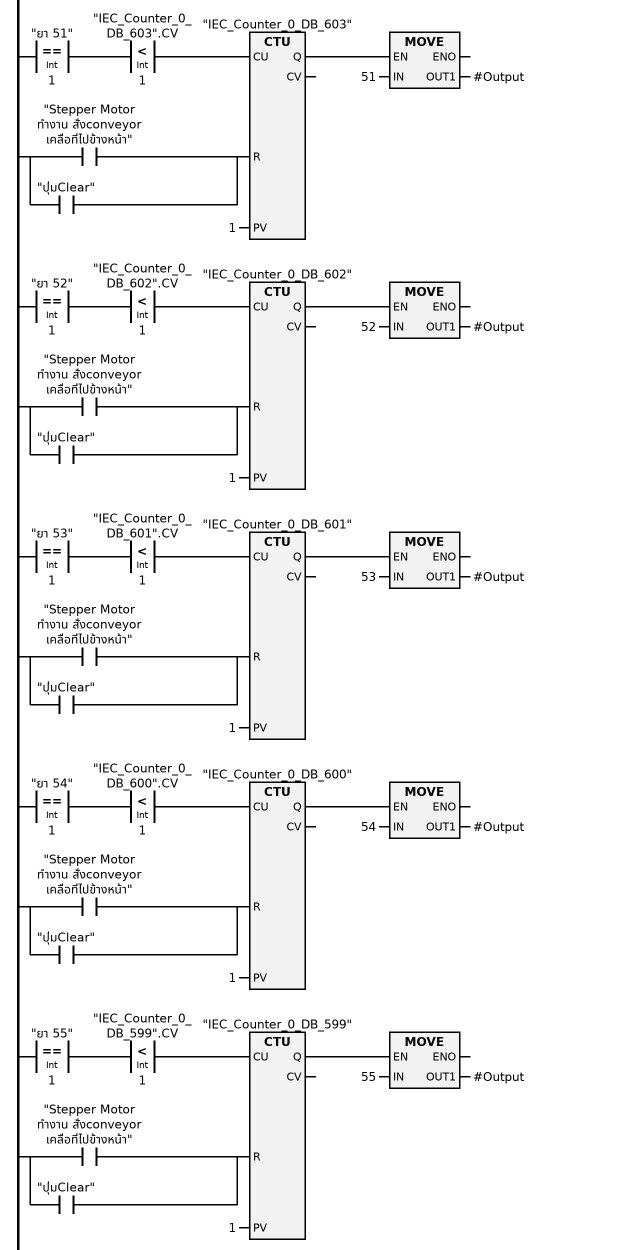
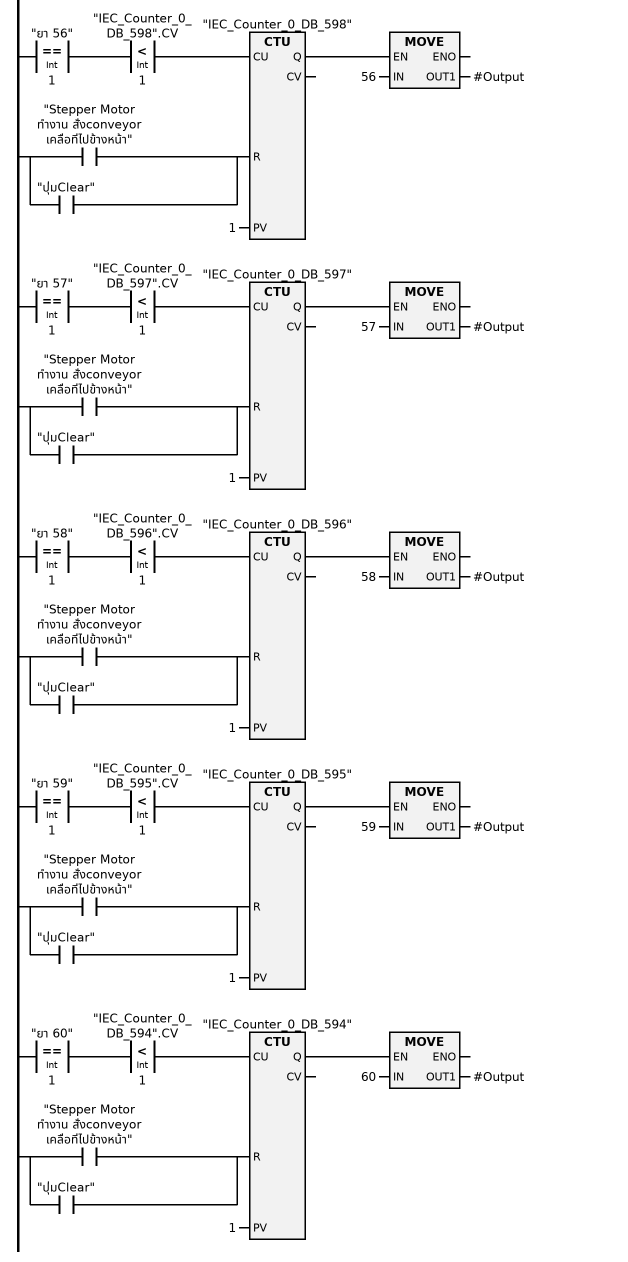
   "IEC_Counter_0_DB_589".CTU(CU := ("ยา 41" = 1) AND ("IEC_Counter_0_DB_589".CV < 1),
                           R := "Stepper Motor ทำงาน สั่งconveyor เคลื่อที่ไปข้างหน้า" OR "ปุ่มClear",
                           PV := 1);
   IF "IEC_Counter_0_DB_589".Q THEN #Output := 41; END_IF;
   "IEC_Counter_0_DB_590".CTU(CU := ("ยา 42" = 1) AND ("IEC_Counter_0_DB_590".CV < 1),
                           R := "Stepper Motor ทำงาน สั่งconveyor เคลื่อที่ไปข้างหน้า" OR "ปุ่มClear",
                           PV := 1);
   IF "IEC_Counter_0_DB_590".Q THEN #Output := 42; END_IF;
   "IEC_Counter_0_DB_591".CTU(CU := ("ยา 43" = 1) AND ("IEC_Counter_0_DB_591".CV < 1),
                           R := "Stepper Motor ทำงาน สั่งconveyor เคลื่อที่ไปข้างหน้า" OR "ปุ่มClear",
                           PV := 1);
   IF "IEC_Counter_0_DB_591".Q THEN #Output := 43; END_IF;
   "IEC_Counter_0_DB_592".CTU(CU := ("ยา 44" = 1) AND ("IEC_Counter_0_DB_592".CV < 1),
                           R := "Stepper Motor ทำงาน สั่งconveyor เคลื่อที่ไปข้างหน้า" OR "ปุ่มClear",
                           PV := 1);
   IF "IEC_Counter_0_DB_592".Q THEN #Output := 44; END_IF;
   "IEC_Counter_0_DB_593".CTU(CU := ("ยา 45" = 1) AND ("IEC_Counter_0_DB_593".CV < 1),
                           R := "Stepper Motor ทำงาน สั่งconveyor เคลื่อที่ไปข้างหน้า" OR "ปุ่มClear",
                           PV := 1);
   IF "IEC_Counter_0_DB_593".Q THEN #Output := 45; END_IF;
   "IEC_Counter_0_DB_608".CTU(CU := ("ยา 46" = 1) AND ("IEC_Counter_0_DB_608".CV < 1),
                           R := "Stepper Motor ทำงาน สั่งconveyor เคลื่อที่ไปข้างหน้า" OR "ปุ่มClear",
                           PV := 1);
   IF "IEC_Counter_0_DB_608".Q THEN #Output := 46; END_IF;
   "IEC_Counter_0_DB_607".CTU(CU := ("ยา 47" = 1) AND ("IEC_Counter_0_DB_607".CV < 1),
                           R := "Stepper Motor ทำงาน สั่งconveyor เคลื่อที่ไปข้างหน้า" OR "ปุ่มClear",
                           PV := 1);
   IF "IEC_Counter_0_DB_607".Q THEN #Output := 47; END_IF;
   "IEC_Counter_0_DB_606".CTU(CU := ("ยา 48" = 1) AND ("IEC_Counter_0_DB_606".CV < 1),
                           R := "Stepper Motor ทำงาน สั่งconveyor เคลื่อที่ไปข้างหน้า" OR "ปุ่มClear",
                           PV := 1);
   IF "IEC_Counter_0_DB_606".Q THEN #Output := 48; END_IF;
   "IEC_Counter_0_DB_605".CTU(CU := ("ยา 49" = 1) AND ("IEC_Counter_0_DB_605".CV < 1),
                           R := "Stepper Motor ทำงาน สั่งconveyor เคลื่อที่ไปข้างหน้า" OR "ปุ่มClear",
                           PV := 1);
   IF "IEC_Counter_0_DB_605".Q THEN #Output := 49; END_IF;
   "IEC_Counter_0_DB_604".CTU(CU := ("ยา 50" = 1) AND ("IEC_Counter_0_DB_604".CV < 1),
                           R := "Stepper Motor ทำงาน สั่งconveyor เคลื่อที่ไปข้างหน้า" OR "ปุ่มClear",
                           PV := 1);
   IF "IEC_Counter_0_DB_604".Q THEN #Output := 50; END_IF;
   "IEC_Counter_0_DB_603".CTU(CU := ("ยา 51" = 1) AND ("IEC_Counter_0_DB_603".CV < 1),
                           R := "Stepper Motor ทำงาน สั่งconveyor เคลื่อที่ไปข้างหน้า" OR "ปุ่มClear",
                           PV := 1);
   IF "IEC_Counter_0_DB_603".Q THEN #Output := 51; END_IF;
   "IEC_Counter_0_DB_602".CTU(CU := ("ยา 52" = 1) AND ("IEC_Counter_0_DB_602".CV < 1),
                           R := "Stepper Motor ทำงาน สั่งconveyor เคลื่อที่ไปข้างหน้า" OR "ปุ่มClear",
                           PV := 1);
   IF "IEC_Counter_0_DB_602".Q THEN #Output := 52; END_IF;
   "IEC_Counter_0_DB_601".CTU(CU := ("ยา 53" = 1) AND ("IEC_Counter_0_DB_601".CV < 1),
                           R := "Stepper Motor ทำงาน สั่งconveyor เคลื่อที่ไปข้างหน้า" OR "ปุ่มClear",
                           PV := 1);
   IF "IEC_Counter_0_DB_601".Q THEN #Output := 53; END_IF;
   "IEC_Counter_0_DB_600".CTU(CU := ("ยา 54" = 1) AND ("IEC_Counter_0_DB_600".CV < 1),
                           R := "Stepper Motor ทำงาน สั่งconveyor เคลื่อที่ไปข้างหน้า" OR "ปุ่มClear",
                           PV := 1);
   IF "IEC_Counter_0_DB_600".Q THEN #Output := 54; END_IF;
   "IEC_Counter_0_DB_599".CTU(CU := ("ยา 55" = 1) AND ("IEC_Counter_0_DB_599".CV < 1),
                           R := "Stepper Motor ทำงาน สั่งconveyor เคลื่อที่ไปข้างหน้า" OR "ปุ่มClear",
                           PV := 1);
   IF "IEC_Counter_0_DB_599".Q THEN #Output := 55; END_IF;
   "IEC_Counter_0_DB_598".CTU(CU := ("ยา 56" = 1) AND ("IEC_Counter_0_DB_598".CV < 1),
                           R := "Stepper Motor ทำงาน สั่งconveyor เคลื่อที่ไปข้างหน้า" OR "ปุ่มClear",
                           PV := 1);
   IF "IEC_Counter_0_DB_598".Q THEN #Output := 56; END_IF;
   "IEC_Counter_0_DB_597".CTU(CU := ("ยา 57" = 1) AND ("IEC_Counter_0_DB_597".CV < 1),
                           R := "Stepper Motor ทำงาน สั่งconveyor เคลื่อที่ไปข้างหน้า" OR "ปุ่มClear",
                           PV := 1);
   IF "IEC_Counter_0_DB_597".Q THEN #Output := 57; END_IF;
   "IEC_Counter_0_DB_596".CTU(CU := ("ยา 58" = 1) AND ("IEC_Counter_0_DB_596".CV < 1),
                           R := "Stepper Motor ทำงาน สั่งconveyor เคลื่อที่ไปข้างหน้า" OR "ปุ่มClear",
                           PV := 1);
   IF "IEC_Counter_0_DB_596".Q THEN #Output := 58; END_IF;
   "IEC_Counter_0_DB_595".CTU(CU := ("ยา 59" = 1) AND ("IEC_Counter_0_DB_595".CV < 1),
                           R := "Stepper Motor ทำงาน สั่งconveyor เคลื่อที่ไปข้างหน้า" OR "ปุ่มClear",
                           PV := 1);
   IF "IEC_Counter_0_DB_595".Q THEN #Output := 59; END_IF;
   "IEC_Counter_0_DB_594".CTU(CU := ("ยา 60" = 1) AND ("IEC_Counter_0_DB_594".CV < 1),
                           R := "Stepper Motor ทำงาน สั่งconveyor เคลื่อที่ไปข้างหน้า" OR "ปุ่มClear",
                           PV := 1);
   IF "IEC_Counter_0_DB_594".Q THEN #Output := 60; END_IF;
END_REGION

REGION Network 4
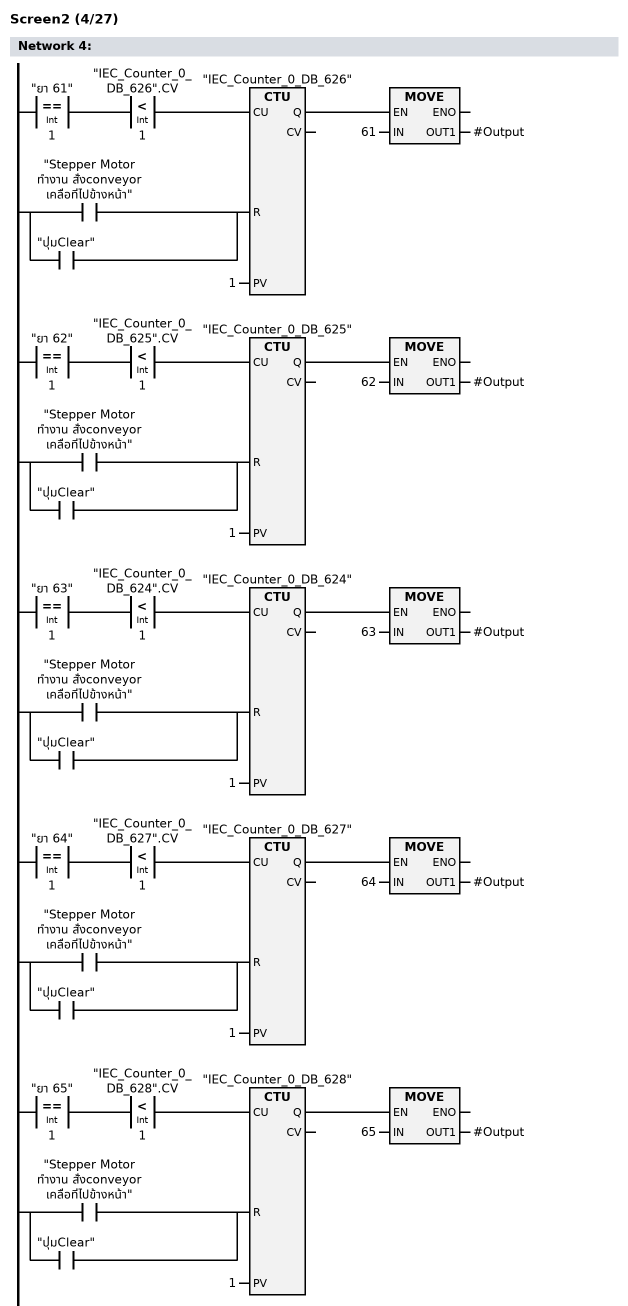
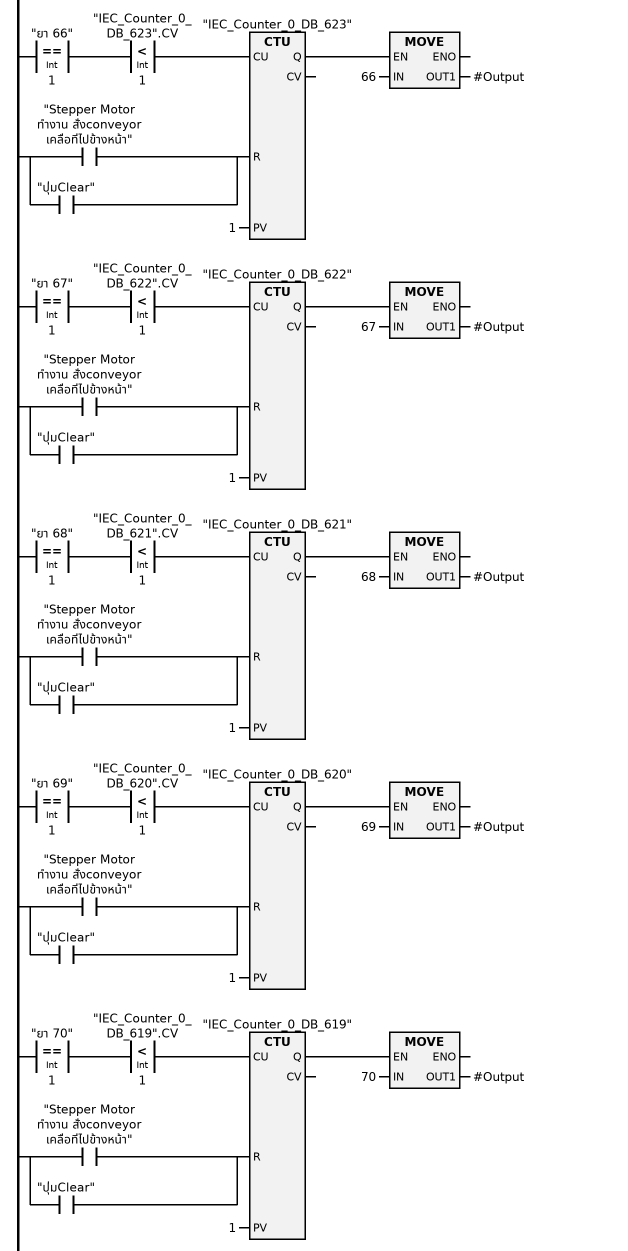
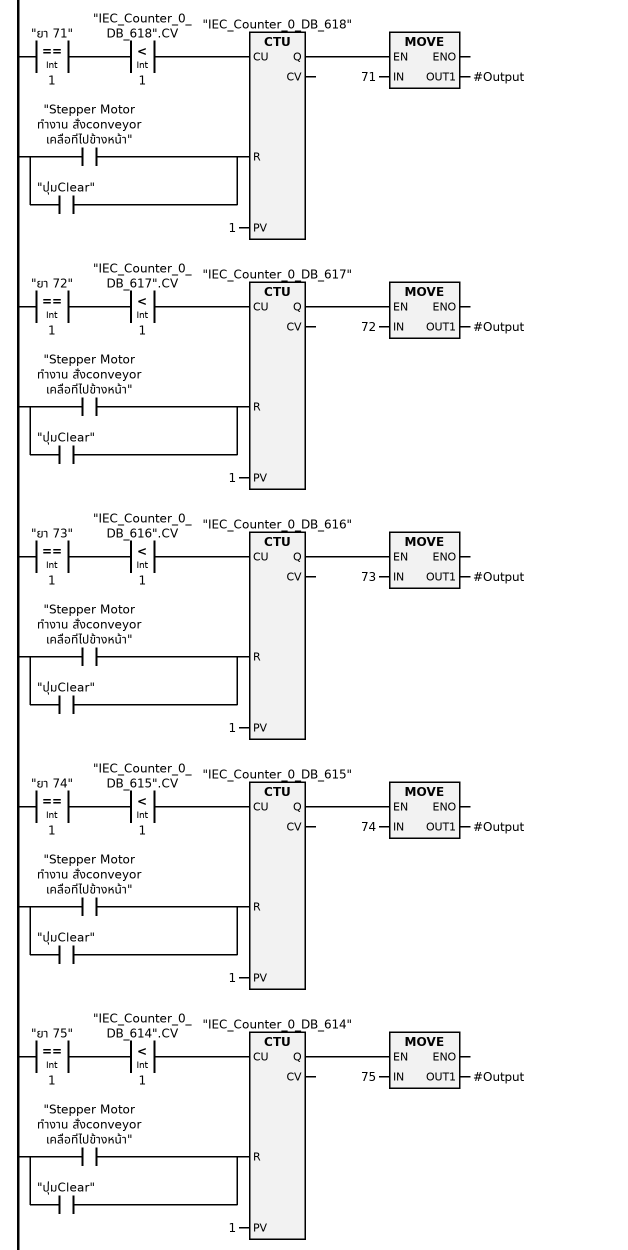
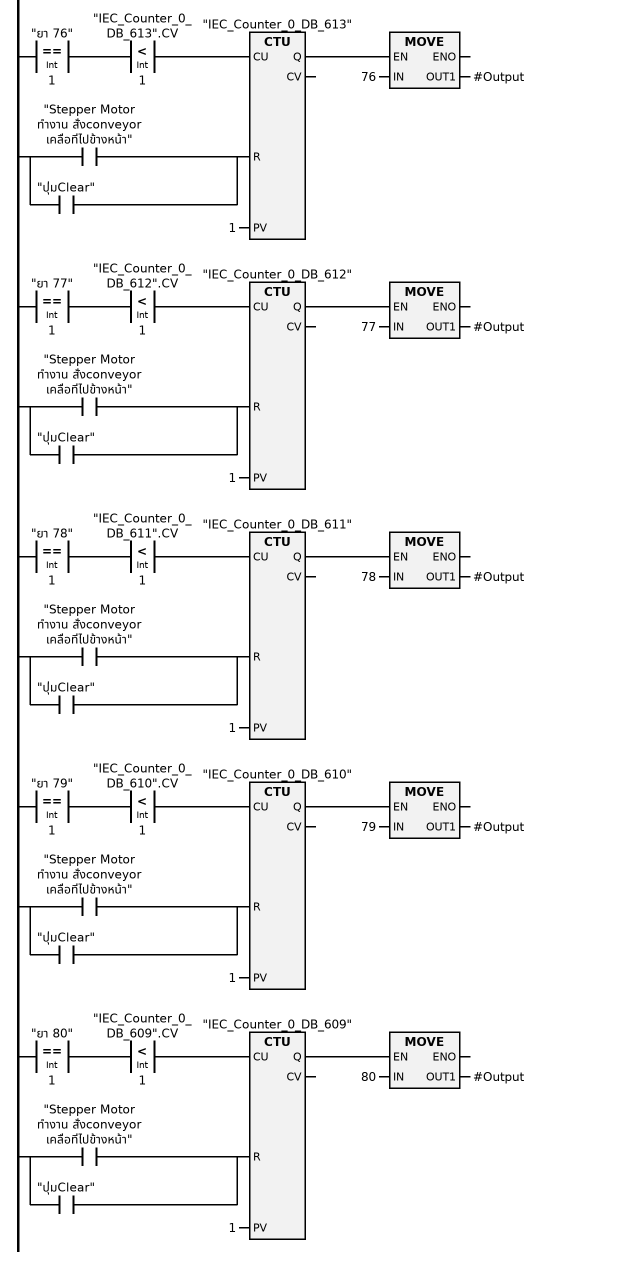
   "IEC_Counter_0_DB_626".CTU(CU := ("ยา 61" = 1) AND ("IEC_Counter_0_DB_626".CV < 1),
                           R := "Stepper Motor ทำงาน สั่งconveyor เคลื่อที่ไปข้างหน้า" OR "ปุ่มClear",
                           PV := 1);
   IF "IEC_Counter_0_DB_626".Q THEN #Output := 61; END_IF;
   "IEC_Counter_0_DB_625".CTU(CU := ("ยา 62" = 1) AND ("IEC_Counter_0_DB_625".CV < 1),
                           R := "Stepper Motor ทำงาน สั่งconveyor เคลื่อที่ไปข้างหน้า" OR "ปุ่มClear",
                           PV := 1);
   IF "IEC_Counter_0_DB_625".Q THEN #Output := 62; END_IF;
   "IEC_Counter_0_DB_624".CTU(CU := ("ยา 63" = 1) AND ("IEC_Counter_0_DB_624".CV < 1),
                           R := "Stepper Motor ทำงาน สั่งconveyor เคลื่อที่ไปข้างหน้า" OR "ปุ่มClear",
                           PV := 1);
   IF "IEC_Counter_0_DB_624".Q THEN #Output := 63; END_IF;
   "IEC_Counter_0_DB_627".CTU(CU := ("ยา 64" = 1) AND ("IEC_Counter_0_DB_627".CV < 1),
                           R := "Stepper Motor ทำงาน สั่งconveyor เคลื่อที่ไปข้างหน้า" OR "ปุ่มClear",
                           PV := 1);
   IF "IEC_Counter_0_DB_627".Q THEN #Output := 64; END_IF;
   "IEC_Counter_0_DB_628".CTU(CU := ("ยา 65" = 1) AND ("IEC_Counter_0_DB_628".CV < 1),
                           R := "Stepper Motor ทำงาน สั่งconveyor เคลื่อที่ไปข้างหน้า" OR "ปุ่มClear",
                           PV := 1);
   IF "IEC_Counter_0_DB_628".Q THEN #Output := 65; END_IF;
   "IEC_Counter_0_DB_623".CTU(CU := ("ยา 66" = 1) AND ("IEC_Counter_0_DB_623".CV < 1),
                           R := "Stepper Motor ทำงาน สั่งconveyor เคลื่อที่ไปข้างหน้า" OR "ปุ่มClear",
                           PV := 1);
   IF "IEC_Counter_0_DB_623".Q THEN #Output := 66; END_IF;
   "IEC_Counter_0_DB_622".CTU(CU := ("ยา 67" = 1) AND ("IEC_Counter_0_DB_622".CV < 1),
                           R := "Stepper Motor ทำงาน สั่งconveyor เคลื่อที่ไปข้างหน้า" OR "ปุ่มClear",
                           PV := 1);
   IF "IEC_Counter_0_DB_622".Q THEN #Output := 67; END_IF;
   "IEC_Counter_0_DB_621".CTU(CU := ("ยา 68" = 1) AND ("IEC_Counter_0_DB_621".CV < 1),
                           R := "Stepper Motor ทำงาน สั่งconveyor เคลื่อที่ไปข้างหน้า" OR "ปุ่มClear",
                           PV := 1);
   IF "IEC_Counter_0_DB_621".Q THEN #Output := 68; END_IF;
   "IEC_Counter_0_DB_620".CTU(CU := ("ยา 69" = 1) AND ("IEC_Counter_0_DB_620".CV < 1),
                           R := "Stepper Motor ทำงาน สั่งconveyor เคลื่อที่ไปข้างหน้า" OR "ปุ่มClear",
                           PV := 1);
   IF "IEC_Counter_0_DB_620".Q THEN #Output := 69; END_IF;
   "IEC_Counter_0_DB_619".CTU(CU := ("ยา 70" = 1) AND ("IEC_Counter_0_DB_619".CV < 1),
                           R := "Stepper Motor ทำงาน สั่งconveyor เคลื่อที่ไปข้างหน้า" OR "ปุ่มClear",
                           PV := 1);
   IF "IEC_Counter_0_DB_619".Q THEN #Output := 70; END_IF;
   "IEC_Counter_0_DB_618".CTU(CU := ("ยา 71" = 1) AND ("IEC_Counter_0_DB_618".CV < 1),
                           R := "Stepper Motor ทำงาน สั่งconveyor เคลื่อที่ไปข้างหน้า" OR "ปุ่มClear",
                           PV := 1);
   IF "IEC_Counter_0_DB_618".Q THEN #Output := 71; END_IF;
   "IEC_Counter_0_DB_617".CTU(CU := ("ยา 72" = 1) AND ("IEC_Counter_0_DB_617".CV < 1),
                           R := "Stepper Motor ทำงาน สั่งconveyor เคลื่อที่ไปข้างหน้า" OR "ปุ่มClear",
                           PV := 1);
   IF "IEC_Counter_0_DB_617".Q THEN #Output := 72; END_IF;
   "IEC_Counter_0_DB_616".CTU(CU := ("ยา 73" = 1) AND ("IEC_Counter_0_DB_616".CV < 1),
                           R := "Stepper Motor ทำงาน สั่งconveyor เคลื่อที่ไปข้างหน้า" OR "ปุ่มClear",
                           PV := 1);
   IF "IEC_Counter_0_DB_616".Q THEN #Output := 73; END_IF;
   "IEC_Counter_0_DB_615".CTU(CU := ("ยา 74" = 1) AND ("IEC_Counter_0_DB_615".CV < 1),
                           R := "Stepper Motor ทำงาน สั่งconveyor เคลื่อที่ไปข้างหน้า" OR "ปุ่มClear",
                           PV := 1);
   IF "IEC_Counter_0_DB_615".Q THEN #Output := 74; END_IF;
   "IEC_Counter_0_DB_614".CTU(CU := ("ยา 75" = 1) AND ("IEC_Counter_0_DB_614".CV < 1),
                           R := "Stepper Motor ทำงาน สั่งconveyor เคลื่อที่ไปข้างหน้า" OR "ปุ่มClear",
                           PV := 1);
   IF "IEC_Counter_0_DB_614".Q THEN #Output := 75; END_IF;
   "IEC_Counter_0_DB_613".CTU(CU := ("ยา 76" = 1) AND ("IEC_Counter_0_DB_613".CV < 1),
                           R := "Stepper Motor ทำงาน สั่งconveyor เคลื่อที่ไปข้างหน้า" OR "ปุ่มClear",
                           PV := 1);
   IF "IEC_Counter_0_DB_613".Q THEN #Output := 76; END_IF;
   "IEC_Counter_0_DB_612".CTU(CU := ("ยา 77" = 1) AND ("IEC_Counter_0_DB_612".CV < 1),
                           R := "Stepper Motor ทำงาน สั่งconveyor เคลื่อที่ไปข้างหน้า" OR "ปุ่มClear",
                           PV := 1);
   IF "IEC_Counter_0_DB_612".Q THEN #Output := 77; END_IF;
   "IEC_Counter_0_DB_611".CTU(CU := ("ยา 78" = 1) AND ("IEC_Counter_0_DB_611".CV < 1),
                           R := "Stepper Motor ทำงาน สั่งconveyor เคลื่อที่ไปข้างหน้า" OR "ปุ่มClear",
                           PV := 1);
   IF "IEC_Counter_0_DB_611".Q THEN #Output := 78; END_IF;
   "IEC_Counter_0_DB_610".CTU(CU := ("ยา 79" = 1) AND ("IEC_Counter_0_DB_610".CV < 1),
                           R := "Stepper Motor ทำงาน สั่งconveyor เคลื่อที่ไปข้างหน้า" OR "ปุ่มClear",
                           PV := 1);
   IF "IEC_Counter_0_DB_610".Q THEN #Output := 79; END_IF;
   "IEC_Counter_0_DB_609".CTU(CU := ("ยา 80" = 1) AND ("IEC_Counter_0_DB_609".CV < 1),
                           R := "Stepper Motor ทำงาน สั่งconveyor เคลื่อที่ไปข้างหน้า" OR "ปุ่มClear",
                           PV := 1);
   IF "IEC_Counter_0_DB_609".Q THEN #Output := 80; END_IF;
END_REGION

REGION Network 5
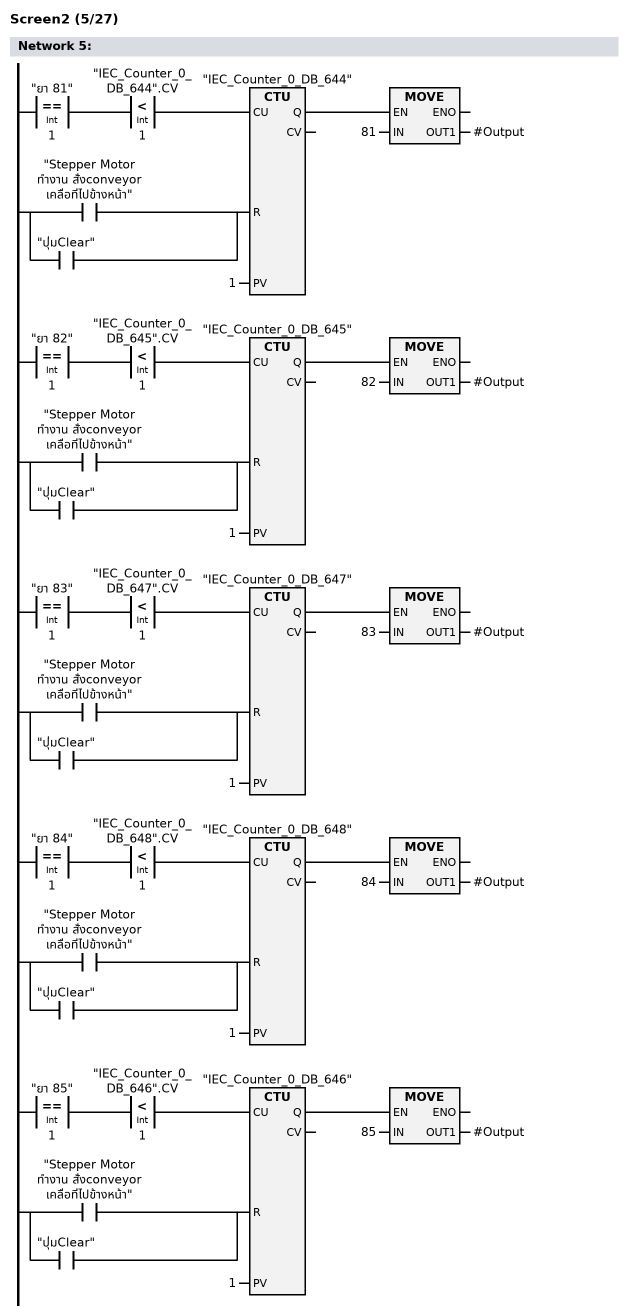
